(* IEC 61131-3 sources: volt/packages/volt-lsp-iec/test-corpus/pro2193/Device/Plc Logic/Application/09 Misc/Library Manager/AlarmManager (part 3) *)

(* ---- ALARMSTORAGEMANAGER.pou ---- *)
FUNCTION_BLOCK ALARMSTORAGEMANAGER
VAR
	M_ALARMSTORAGE : STI.Storage;
	M_ITFSTORAGE : STO.IStorage;
	M_ITFTABLE : STO.ITable;
	M_ADWROOTPAGES : ARRAY [EAlarmStorageObject.IX_MIN..EAlarmStorageObject.IX_LAST] OF CAA.IDENT;
	M_XROOTPAGESDETERMINED : BOOL;
	M_UDICOUNTLATCHVARIABLES : CAA.COUNT;
	WRITEACCESSNECESSARY : BOOL;
END_VAR
END_FUNCTION_BLOCK

METHOD BEGINTRANSACTION : STO.ITransaction
VAR_INPUT
	XREADONLY : BOOL;
END_VAR
VAR_OUTPUT
	EERROR : STO.ERROR;
END_VAR
END_METHOD

METHOD CLOSETABLE
VAR_INPUT
	ITFTABLE : STO.ITable;
END_VAR
END_METHOD

METHOD ENDTRANSACTION
VAR_INPUT
	ITFTRANSACTION : STO.ITransaction;
	EERROR : STO.ERROR;
END_VAR
END_METHOD

METHOD FB_EXIT : BOOL
VAR_INPUT
	BINCOPYCODE : BOOL;
END_VAR
END_METHOD

METHOD GETCOLUMNIDENTIFIER : CAA.IDENT
VAR_INPUT
	IDCOLUMN : CAA.IDENT;
END_VAR
END_METHOD

METHOD GETNUMBEROFLATCHVARIABLES : CAA.COUNT
VAR_INPUT
	IDBVERSION : INT;
	UDICOUNTCOLUMNSTBLALARM : CAA.COUNT;
END_VAR
END_METHOD

METHOD GETSTORAGE : STO.IStorage
END_METHOD

METHOD OPENTABLE : STO.ITable
VAR_INPUT
	XREADONLY : BOOL;
END_VAR
VAR_OUTPUT
	EERROR : STO.ERROR;
END_VAR
END_METHOD

METHOD DETERMINEROOTPAGES : STO.ERROR
END_METHOD

METHOD GETROOTPAGE : CAA.IDENT
VAR_INPUT
	EDATABASEOBJECT : EAlarmStorageObject;
END_VAR
END_METHOD

METHOD ISREADY : BOOL
END_METHOD

METHOD RESET
END_METHOD

METHOD CLOSESTORAGE
END_METHOD

METHOD DETERMINEROOTPAGESOPENSTORAGE : STO.ERROR
VAR_OUTPUT
	XREOPENREADONLY : BOOL;
END_VAR
END_METHOD

METHOD PRVCHECKJOURNAL
END_METHOD

METHOD PRVHELPGETDATABASEFILEPATH : CAA.FILENAME
END_METHOD

METHOD PRVOPENSTORAGE : STO.ERROR
VAR_INPUT
	XREADONLY : BOOL;
END_VAR
END_METHOD

METHOD PROTCLOSECURSOR : STO.ERROR
VAR_INPUT
	EERRORFROMPREVIOUSPROCESSING : STO.ERROR;
	ICALLINGMETHOD : INT;
END_VAR
VAR_IN_OUT
	ITFCURSOR : STO.ICursor;
END_VAR
END_METHOD

METHOD PROTGETEXCLUSIVETRANSACTION : STO.ITransaction
VAR_INPUT
	ICOUNTRETRIES : INT;
END_VAR
VAR_OUTPUT
	EERROR : STO.ERROR;
END_VAR
END_METHOD

METHOD PROTRELEASEROW : STO.ERROR
VAR_INPUT
	EERRORFROMPREVIOUSPROCESSING : STO.ERROR;
	ICALLINGMETHOD : INT;
END_VAR
VAR_IN_OUT
	ITFROW : STO.IRow;
END_VAR
END_METHOD

(* ---- ALARMSTORAGEQUEUE.pou ---- *)
FUNCTION_BLOCK ALARMSTORAGEQUEUE
VAR
	_PAQUEUE : POINTER TO ARRAY [0..0] OF AlarmStorageRow;
	_IQUEUESIZE : UDINT;
	_INEWESTPOS : UDINT := 0;
	_IOLDESTPOS : UDINT := 0;
	_IITEMCOUNT : UDINT := 0;
	_ALARMSTORAGEROWPROVIDER : AlarmStorageRowProvider;
	_UICOUNTEVENTS : UDINT;
	_PAINITIALQUEUE : POINTER TO AlarmStorageRow;
	_XKEEPOLDVALUES : BOOL;
	_XFIXQUEUENECESSARY : BOOL;
	COUNTALARMSTOINSERT : UDINT;
	COUNTEVENTSTOINSERT : UDINT;
END_VAR
END_FUNCTION_BLOCK

METHOD CANPOSTALARM : BOOL
END_METHOD

METHOD CLEAR
END_METHOD

METHOD FB_EXIT : BOOL
VAR_INPUT
	BINCOPYCODE : BOOL;
END_VAR
END_METHOD

METHOD FB_INIT : BOOL
VAR_INPUT
	BINITRETAINS : BOOL;
	BINCOPYCODE : BOOL;
END_VAR
END_METHOD

METHOD FIXAFTERONLINECHANGEIFNECESSARY
VAR_INPUT
	STORAGE : IDatabaseFileAlarmStorage;
END_VAR
END_METHOD

METHOD GETCURRENTALARM : AlarmStorageRow
END_METHOD

METHOD INIT
VAR_INPUT
	PQUEUEDATA : POINTER TO AlarmStorageRow;
	NUMQUEUEENTRIES : UDINT;
END_VAR
END_METHOD

METHOD ISEMPTY : BOOL
END_METHOD

METHOD ONLINECHANGEDONE
END_METHOD

METHOD ONLINECHANGEPREPARE
END_METHOD

METHOD POSTALARM : BOOL
VAR_INPUT
	ITFALARM : IAlarm;
	ITFDATABASEFILEALARMSTORAGE : IDatabaseFileAlarmStorage;
	ESTATE : AlarmState;
	EPREVSTATE : AlarmState;
	XFORCEUPDATE : BOOL;
END_VAR
VAR_OUTPUT
	ROW : AlarmStorageRow;
END_VAR
END_METHOD

METHOD REMOVECURRENTALARM
END_METHOD

METHOD TRYTOENLARGEQUEUE
END_METHOD

METHOD ASSIGNINITVALUES
END_METHOD

METHOD RESETSTOREDREFERENCES
END_METHOD

METHOD TRYTOENLARGEQUEUEHELP
VAR_INPUT
	KEEPNEWESTPOS : BOOL;
END_VAR
END_METHOD

METHOD PRVGETTYPEDVALUE
VAR_INPUT
	ITFTYPEDVALUE : ITypedValue;
END_VAR
VAR_OUTPUT
	BYTYPECLASS : BYTE;
	LIVALUE : LINT;
END_VAR
END_METHOD

(* ---- ALARMSTORAGEREADER.pou ---- *)
FUNCTION_BLOCK ALARMSTORAGEREADER EXTENDS AlarmStorageManager
VAR_INPUT
	_HLOCK : RTS_IEC_HANDLE := RTS_INVALID_HANDLE;
END_VAR
VAR
	M_DATABASEACCESS : SQLiteDatabaseAccess;
	M_ROWIDITERATOR : AlarmStorageReaderRowIdIterator;
	M_ITFALARMSTORAGEREADERCONSUMER : IAlarmStorageReaderConsumer;
	M_ITFALARMSTORAGEMANAGER : IAlarmStorageManager := THIS^;
	M_EBYTEORDER : EAlarmByteOrder := EAlarmByteOrder.Unknown;
	M_ALATCHVARIABLES : ARRAY [1..2] OF LatchVariable;
	M_AWSLATCHVARVALUE : ARRAY [0..1] OF WSTRING(255);
	M_PALATCHVARSTRINGALLOC : POINTER TO ARRAY [0..10] OF WSTRING(255);
	M_PALATCHVARALLOC : POINTER TO ARRAY [0..10] OF LatchVariable;
	M_ICOUNTLATCHVARALLOC : INT;
	M_LOCKRESULT : RTS_IEC_RESULT;
	M_SWHOHASLOCK : STRING;
END_VAR
END_FUNCTION_BLOCK

METHOD ADDALARMSTORAGELISTENER : EAlarmStorageReaderErrors
VAR_INPUT
	ITFALARMSTORAGELISTENER : IAlarmStorageListener;
END_VAR
END_METHOD

METHOD CONTINUEREADING : EAlarmStorageReaderErrors
VAR_INPUT
	LITIMSTAMPFROM : LINT;
	LITIMSTAMPTO : LINT;
	XREADASCENDING : BOOL;
	ITFALARMSTORAGEREADERCONSUMER : IAlarmStorageReaderConsumer;
END_VAR
END_METHOD

METHOD FB_EXIT : BOOL
VAR_INPUT
	BINCOPYCODE : BOOL;
END_VAR
END_METHOD

METHOD FB_INIT : BOOL
VAR_INPUT
	BINITRETAINS : BOOL;
	BINCOPYCODE : BOOL;
END_VAR
END_METHOD

METHOD GETALARMSFROMSTORAGE : STO.ERROR
VAR_INPUT
	ISKIPROWS : INT;
	IMAXROWS : INT;
	FILTERCRITERIA : REFERENCE TO VisuFbAlarmFilterCriteria;
	ITFALARMDATABLOCK : IAlarmDataBlockBase2;
END_VAR
VAR_IN_OUT
	BROWIDVALID : BOOL;
	DIROWID : DINT;
END_VAR
END_METHOD

METHOD GETALARMSFROMSTORAGE2 : STO.ERROR
VAR_INPUT
	ITFDATABASEACCESS : IDatabaseAccess;
	ISKIPROWS : INT;
	IMAXROWS : INT;
	FILTERCRITERIA : REFERENCE TO VisuFbAlarmFilterCriteria;
	ITFALARMDATABLOCK : IAlarmDataBlockBase2;
END_VAR
VAR_IN_OUT
	BROWIDVALID : BOOL;
	DIROWID : DINT;
END_VAR
END_METHOD

METHOD GETALARMSFROMSTORAGE3 : STO.ERROR
VAR_INPUT
	ITFDATABASEACCESS : IDatabaseAccess3;
	DWROWIDLATEST : DWORD;
	IMAXROWS : INT;
	ITFALARMTRAVERSALCONSUMER : IAlarmTraversalConsumer;
END_VAR
END_METHOD

METHOD GETALARMSFROMSTORAGE4 : STO.ERROR
VAR_INPUT
	ITFDATABASEACCESS : IDatabaseAccess3;
	ITFALARMTRAVERSALCONSUMER : IAlarmTraversalConsumer;
END_VAR
END_METHOD

METHOD GETALARMSFROMSTORAGE5 : STO.ERROR
VAR_INPUT
	DISKIPROWS : DINT;
	DIMAXROWS : DINT;
	FILTERCRITERIA : REFERENCE TO VisuFbAlarmFilterCriteria;
	ITFALARMDATABLOCK : IAlarmDataBlockBase2;
END_VAR
VAR_IN_OUT
	BROWIDVALID : BOOL;
	DIROWID : DINT;
END_VAR
END_METHOD

METHOD GETALARMSFROMSTORAGE6 : STO.ERROR
VAR_INPUT
	ITFDATABASEACCESS : IDatabaseAccess;
	DISKIPROWS : DINT;
	DIMAXROWS : DINT;
	FILTERCRITERIA : REFERENCE TO VisuFbAlarmFilterCriteria;
	ITFALARMDATABLOCK : IAlarmDataBlockBase2;
END_VAR
VAR_IN_OUT
	BROWIDVALID : BOOL;
	DIROWID : DINT;
END_VAR
END_METHOD

METHOD GETCOUNTALARMSFROMSTORAGE : DINT
VAR_INPUT
	FILTERCRITERIA : REFERENCE TO VisuFbAlarmFilterCriteria;
	ITFALARMDATABLOCK : IAlarmDataBlockBase2;
END_VAR
VAR_OUTPUT
	EERROR : STO.ERROR;
	DWCOUNTLATCHVARIABLESINSTORAGE : CAA.COUNT;
END_VAR
END_METHOD

METHOD GETCOUNTALLALARMSFROMSTORAGE : CAA.COUNT
VAR_OUTPUT
	EERROR : STO.ERROR;
END_VAR
END_METHOD

METHOD GETFIRSTLASTROWID : EAlarmStorageReaderErrors
VAR_OUTPUT
	DIROWIDFIRST : DINT;
	DIROWIDLAST : DINT;
END_VAR
END_METHOD

METHOD GETMINMAXTIMESTAMPS : EAlarmStorageReaderErrors
VAR_OUTPUT
	LIMINTIMESTAMP : LINT;
	LIMAXTIMESTAMP : LINT;
	XTABLEISEMPTY : BOOL;
	UDICOUNTALARMS : UDINT;
END_VAR
END_METHOD

METHOD READ : EAlarmStorageReaderErrors
VAR_INPUT
	LITIMSTAMPFROM : LINT;
	LITIMSTAMPTO : LINT;
	XREADASCENDING : BOOL;
	ITFALARMSTORAGEREADERCONSUMER : IAlarmStorageReaderConsumer;
END_VAR
END_METHOD

METHOD REMOVEALARMSTORAGELISTENER : EAlarmStorageReaderErrors
VAR_INPUT
	ITFALARMSTORAGELISTENER : IAlarmStorageListener;
END_VAR
END_METHOD

METHOD SEMAPHOREACQUIRE
VAR_INPUT
	SWHO : STRING;
END_VAR
END_METHOD

METHOD SEMAPHORERELEASE
VAR_INPUT
	SWHO : STRING;
END_VAR
END_METHOD

METHOD PRVALLOCLATCHVARS
VAR_INPUT
	ICNTVAR : INT;
END_VAR
END_METHOD

METHOD PRVDOCONTINUEREADING : BOOL
VAR_INPUT
	DIROWCOUNTER : DINT;
END_VAR
END_METHOD

METHOD PRVFINDROWID : CAA.IDENT
VAR_INPUT
	ITFDATABASEACCESS : IDatabaseAccess;
	XSEARCHFIRST : BOOL;
END_VAR
VAR_OUTPUT
	EERROR : STO.ERROR;
END_VAR
END_METHOD

METHOD PRVFREELATCHVARS
END_METHOD

METHOD PRVREAD : EAlarmStorageReaderErrors
VAR_INPUT
	LITIMSTAMPFROM : LINT;
	LITIMSTAMPTO : LINT;
	XREADASCENDING : BOOL;
END_VAR
END_METHOD

METHOD PRVREADALARMCOMMENT
VAR_INPUT
	IDWHICHCOLUMN : CAA.IDENT;
	ITFDATABASEACCESS4 : IDatabaseAccess4;
END_VAR
VAR_IN_OUT
	EERROR : STO.ERROR;
	CMTBUFFER : AlarmComment;
END_VAR
END_METHOD

METHOD PRVREADLATCHVARSTRING2 : STO.ERROR
VAR_INPUT
	LIROWID : LINT;
	ITFDATABASEACCESS : IDatabaseAccess;
	BYLATCHVARTYPE : BYTE;
	PBVARVALUE : POINTER TO BYTE;
	ISZVARVALUE : INT;
END_VAR
END_METHOD

METHOD PRVREADLATCHVARSTRING : STO.ERROR
VAR_INPUT
	LIROWID : LINT;
	ITFDATABASEACCESS : IDatabaseAccess;
	BYLATCHVARTYPE : BYTE;
END_VAR
VAR_OUTPUT
	CBPSTRING : CharBufferPtr;
END_VAR
END_METHOD

METHOD PRVRETRIEVELATCHVARVALUE : STO.ERROR
VAR_INPUT
	ITFDATABASEACCESS : IDatabaseAccess;
	ITFALARMMETAOBJECTSTUB3 : IAlarmMetaObjectStub3;
	USIWHICHLATCHVAR : USINT;
END_VAR
END_METHOD

METHOD PRVTBLALARMFINDTIMESTAMP : STO.ERROR
VAR_INPUT
	ITFDATABASEACCESS : IDatabaseAccess;
	LITIMSTAMP : LINT;
	XUSENEXTROW : BOOL;
END_VAR
VAR_OUTPUT
	IDROWTIMSTAMP : CAA.IDENT;
END_VAR
END_METHOD

(* ---- ALARMSTORAGEREADERROWIDITERATOR.pou ---- *)
FUNCTION_BLOCK ALARMSTORAGEREADERROWIDITERATOR
VAR
	M_IDROWTBLALARMFROM : CAA.IDENT;
	M_IDROWTBLALARMTO : CAA.IDENT;
	M_IDROWCURR : CAA.IDENT;
	M_XITERATEASCENDING : BOOL;
	M_IDLASTPROCESSEDROWID : CAA.IDENT := AlarmConstants.INVALID_ROWID;
	M_LITIMESTAMP : LINT;
END_VAR
END_FUNCTION_BLOCK

METHOD GETNEXTROWID : CAA.IDENT
END_METHOD

METHOD GETSAVEDSTATE : LINT
END_METHOD

METHOD HASNEXTROWID : BOOL
END_METHOD

METHOD HASSAVEDSTATE : BOOL
END_METHOD

METHOD INITIALIZE
VAR_INPUT
	IDROWTBLALARMFROM : CAA.IDENT;
	IDROWTBLALARMTO : CAA.IDENT;
	XITERATEASCENDING : BOOL;
END_VAR
END_METHOD

METHOD SAVESTATE
VAR_INPUT
	IDLASTPROCESSEDROWID : CAA.IDENT;
	LITIMESTAMP : LINT;
END_VAR
END_METHOD

(* ---- ALARMSTORAGEROW.pou ---- *)
FUNCTION_BLOCK ALARMSTORAGEROW
VAR_INPUT
	UDIALARMID : UDINT;
	UDIALARMCLASSID : UDINT;
	UDIALARMGROUPID : UDINT;
	LITIMESTAPLAST : TIMESTAMP;
	LITIMESTAPACTIVE : TIMESTAMP;
	LITIMESTAPINACTIVE : TIMESTAMP;
	LITIMESTAPACKNOWLEDGE : TIMESTAMP;
	IOFFSETLAST : INT := -1;
	IOFFSETACTIVE : INT := -1;
	IOFFSETINACTIVE : INT := -1;
	IOFFSETACKNOWLEDGE : INT := -1;
	USIPRIORITY : USINT;
	ESTATE : AlarmState;
	EPREVSTATE : AlarmState;
	BYTRIGGERVALUETYPE : BYTE;
	LITRIGGERVALUEVAL : LINT;
	PLATCHVARIABLES : POINTER TO ARRAY [0..10] OF LatchVariable;
	USICOUNTLATCHVARIABLES : USINT;
	ITFALARM : IAlarm;
	ITFDATABASEFILEALARMSTORAGE : IDatabaseFileAlarmStorage;
	IDROW : CAA.IDENT;
	XIDROWVALID : BOOL;
	XFORCEUPDATE : BOOL;
	SREMOTEDEVICENAME : STRING;
	CMTACTIVE : AlarmComment;
	CMTACTIVEACK : AlarmComment;
	CMTWAITINGCONF : AlarmComment;
	CMTNORMAL : AlarmComment;
	XINVALID : BOOL;
END_VAR
END_FUNCTION_BLOCK

METHOD DERIVEALARMREFERENCE
END_METHOD

METHOD GETLATCHVARVALUE
VAR_INPUT
	USIWHICHLATCHVAR : USINT;
END_VAR
VAR_OUTPUT
	BYTYPE : BYTE;
	LIVALUE : LINT;
END_VAR
END_METHOD

METHOD RESETALARMCOMMENTS : BOOL
END_METHOD

METHOD SETLATCHVARVALUE
VAR_INPUT
	USIWHICHLATCHVAR : USINT;
	BYTYPE : BYTE;
	LIVALUE : LINT;
END_VAR
END_METHOD

(* ---- ALARMSTORAGEROWPROVIDER.pou ---- *)
FUNCTION_BLOCK ALARMSTORAGEROWPROVIDER
VAR
	M_PAALARMSTORAGEROWS : POINTER TO ARRAY [0..100] OF AlarmStorageRow;
	M_ICOUNTROWS : UDINT;
	M_PALATCHVARIABLES : POINTER TO ARRAY [0..100] OF LatchVariable;
	M_ICOUNTLATCHVARIABLES : UDINT;
	COMPONENT : STRING := 'AlarmStorageRowProvider';
END_VAR
END_FUNCTION_BLOCK

METHOD ALLOCATEALARMSTORAGEROWARRAY : BOOL
VAR_INPUT
	IREQUIREDARRAYSIZE : UDINT;
	USICOUNTLATCHVARIABLES : USINT;
	PACURRENTQUEUE : POINTER TO AlarmStorageRow;
	ICURRENTQUEUESIZE : UDINT;
	ICURRENTREADINDEX : UDINT;
END_VAR
VAR_OUTPUT
	PANEWQUEUE : POINTER TO ARRAY [0..0] OF AlarmStorageRow;
	INEWQUEUESIZE : UDINT;
END_VAR
END_METHOD

METHOD COPYQUEUECONTENT : BOOL
VAR_INPUT
	PACURRENTQUEUE : POINTER TO AlarmStorageRow;
	ICURRENTQUEUESIZE : UDINT;
	ICURRENTREADINDEX : UDINT;
	PANEWALARMSTORAGEROWS : POINTER TO AlarmStorageRow;
	INEWQUEUESIZE : UDINT;
	PANEWLATCHVARIABLES : POINTER TO LatchVariable;
	USICOUNTLATCHVARIABLES : USINT;
END_VAR
END_METHOD

METHOD FB_EXIT : BOOL
VAR_INPUT
	BINCOPYCODE : BOOL;
END_VAR
END_METHOD

METHOD FREEBUFFER
VAR_INPUT
	PPBYBUFFER : POINTER TO POINTER TO BYTE;
	PICOUNT : POINTER TO INT;
END_VAR
END_METHOD

METHOD FREEBUFFERS
END_METHOD

(* ---- ALLOCATOR.pou ---- *)
FUNCTION_BLOCK ALLOCATOR
VAR_INPUT
	SCOMPONENT : STRING;
END_VAR
VAR
	DITOTMEM : DINT;
	TOTMEM : DINT;
END_VAR
END_FUNCTION_BLOCK

METHOD ALLOCANDCOPYWSTRING : POINTER TO WSTRING
VAR_INPUT
	PWSWHO : POINTER TO WSTRING;
END_VAR
END_METHOD

METHOD ALLOCBYTES : POINTER TO BYTE
VAR_INPUT
	UXISIZE : __UXINT;
	SWHO : STRING;
END_VAR
END_METHOD

METHOD ALLOCPROXYFBALARMCONTAINER : POINTER TO AlarmContainer
VAR_INPUT
	SWHO : STRING;
END_VAR
END_METHOD

METHOD ALLOCPROXYFBALARMMETAOBJECTSTUB : POINTER TO ProxyFbAlarmMetaObjectStub
VAR_INPUT
	SWHO : STRING;
END_VAR
END_METHOD

METHOD ALLOCPROXYSTRUCTALARMCLASSDESCRIPTION : POINTER TO ProxyStructAlarmClass
VAR_INPUT
	SWHO : STRING;
END_VAR
END_METHOD

METHOD ALLOCPROXYSTRUCTALARMDESCRIPTION : POINTER TO ProxyStructAlarm
VAR_INPUT
	SWHO : STRING;
END_VAR
END_METHOD

METHOD ALLOCPROXYSTRUCTALARMGROUPDESCRIPTION : POINTER TO ProxyStructAlarmGroup
VAR_INPUT
	SWHO : STRING;
END_VAR
END_METHOD

METHOD ALLOCPROXYSTRUCTHISTORICALALARMACTIVE : POINTER TO ProxyStructHistoricalAlarmActive
VAR_INPUT
	SWHO : STRING;
END_VAR
END_METHOD

METHOD ALLOCVALUETYPEBUNDLE : POINTER TO ValueTypeBundle
VAR_INPUT
	SWHO : STRING;
END_VAR
END_METHOD

METHOD FREEBYTES
VAR_INPUT
	PTR : POINTER TO BYTE;
	UXISIZE : __UXINT;
END_VAR
END_METHOD

METHOD FREEPROXYFBALARMCONTAINER
VAR_INPUT
	PREQ : POINTER TO AlarmContainer;
END_VAR
END_METHOD

METHOD FREEPROXYFBALARMMETAOBJECTSTUB
VAR_INPUT
	PREQ : POINTER TO ProxyFbAlarmMetaObjectStub;
END_VAR
END_METHOD

METHOD FREEPROXYSTRUCTALARMCLASSDESCRIPTION
VAR_INPUT
	PREQ : POINTER TO ProxyStructAlarmGroup;
END_VAR
END_METHOD

METHOD FREEPROXYSTRUCTALARMDESCRIPTION
VAR_INPUT
	PREQ : POINTER TO ProxyStructAlarm;
END_VAR
END_METHOD

METHOD FREEPROXYSTRUCTALARMGROUPDESCRIPTION
VAR_INPUT
	PREQ : POINTER TO ProxyStructAlarmClass;
END_VAR
END_METHOD

METHOD FREEPROXYSTRUCTHISTORICALALARMACTIVE
VAR_INPUT
	PREQ : POINTER TO ProxyStructHistoricalAlarmActive;
END_VAR
END_METHOD

METHOD FREEVALUETYPEBUNDLE
VAR_INPUT
	PREQ : POINTER TO ValueTypeBundle;
END_VAR
END_METHOD

(* ---- BINTAGWRITERALARMMETAOBJECTSTUB.pou ---- *)
FUNCTION_BLOCK BINTAGWRITERALARMMETAOBJECTSTUB
VAR
	M_ITFTAGGEDSERVICEWRITER : ITaggedServiceWriter;
	M_LITIMESTAMPACKNOWLEDGE : Timestamp;
	M_LITIMESTAMPACTIVE : Timestamp;
	M_LITIMESTAMPINACTIVE : Timestamp;
	M_LITIMESTAMPLAST : Timestamp;
	M_ITFTYPEDVALUETRIGGER : ITypedValue;
	M_IOFFSETACKNOWLEDGE : INT := -1;
	M_IOFFSETACTIVE : INT := -1;
	M_IOFFSETINACTIVE : INT := -1;
	M_IOFFSETLAST : INT := -1;
	M_PALATCHVARIABLES : POINTER TO ARRAY [0..0] OF LatchVariable;
	M_ICOUNTLATCHVARIABLES : INT;
	M_ISTATE : INT;
	M_UDIALARMID : UDINT;
	M_UDIALARMGROUPID : UDINT;
	OFFSETACKNOWLEDGE : INT;
	OFFSETACTIVE : INT;
	OFFSETINACTIVE : INT;
	OFFSETLAST : INT;
END_VAR
END_FUNCTION_BLOCK

METHOD INITIALIZE
VAR_INPUT
	ITFTAGGEDSERVICEWRITER : ITaggedServiceWriter;
END_VAR
END_METHOD

METHOD SETLATCHVARIABLESBUFFER
VAR_INPUT
	PALATCHVARIABLES : POINTER TO ARRAY [0..0] OF LatchVariable;
	ICOUNTLATCHVARIABLES : INT;
END_VAR
END_METHOD

METHOD SETLATCHVAR1VALUE
VAR_INPUT
	ITFTYPEDVALUELATCHVAR1 : ITypedValue;
END_VAR
END_METHOD

METHOD SETLATCHVAR2VALUE
VAR_INPUT
	ITFTYPEDVALUELATCHVAR2 : ITypedValue;
END_VAR
END_METHOD

METHOD SETSTATE
VAR_INPUT
	ISTATE : INT;
END_VAR
END_METHOD

METHOD SETTIMESTAMPACKNOWLEDGE
VAR_INPUT
	LITIMESTAMPACKNOWLEDGE : Timestamp;
END_VAR
END_METHOD

METHOD SETTIMESTAMPACTIVE
VAR_INPUT
	LITIMESTAMPACTIVE : Timestamp;
END_VAR
END_METHOD

METHOD SETTIMESTAMPINACTIVE
VAR_INPUT
	LITIMESTAMPINACTIVE : Timestamp;
END_VAR
END_METHOD

METHOD SETTIMESTAMPLAST
VAR_INPUT
	LITIMESTAMPLAST : Timestamp;
END_VAR
END_METHOD

METHOD SETTRIGGERVALUE
VAR_INPUT
	ITFTYPEDVALUETRIGGER : ITypedValue;
END_VAR
END_METHOD

METHOD GETCOUNTLATCHVARIABLES : USINT
END_METHOD

METHOD GETLATCHVARVALUE : ITypedValue2
VAR_INPUT
	IWHICHLATCHVAR : INT;
END_VAR
END_METHOD

METHOD SETLATCHVARVALUE
VAR_INPUT
	IWHICHLATCHVAR : INT;
	ITFTYPEDVALUELATCHVAR : ITypedValue;
END_VAR
END_METHOD

METHOD SETALARM
VAR_INPUT
	PALARM : POINTER TO Alarm;
END_VAR
END_METHOD

METHOD FILLINGCOMPLETED : UDINT
END_METHOD

METHOD PRVGETTYPE : BYTE
VAR_INPUT
	ITFTYPEDVALUE : ITypedValue;
END_VAR
END_METHOD

METHOD PRVGETVALUE : LWORD
VAR_INPUT
	ITFTYPEDVALUE : ITypedValue;
END_VAR
END_METHOD

METHOD PRVWRITELATCHVARIABLE
VAR_INPUT
	IWHICHLATCHVAR : INT;
END_VAR
END_METHOD

METHOD GETALARMGROUP : STRING
END_METHOD

METHOD GETCHECKSUM : UDINT
END_METHOD

METHOD GETCURRENTVALUE : ITypedValue
END_METHOD

METHOD GETID : ALARM_ID
END_METHOD

METHOD GETLATCHVAR1VALUE : ITypedValue
END_METHOD

METHOD GETLATCHVAR2VALUE : ITypedValue
END_METHOD

METHOD GETSTATE : INT
END_METHOD

METHOD GETTIMESTAMPACKNOWLEDGE : Timestamp
END_METHOD

METHOD GETTIMESTAMPACTIVE : Timestamp
END_METHOD

METHOD GETTIMESTAMPINACTIVE : Timestamp
END_METHOD

METHOD GETTIMESTAMPLAST : Timestamp
END_METHOD

METHOD GETTRIGGERVALUE : ITypedValue
END_METHOD

METHOD SETACKNOWLEDGE
VAR_INPUT
	BACKNOWLEDGEMULTIPLE : BOOL;
END_VAR
END_METHOD

METHOD SETALARMGROUP
VAR_INPUT
	SALARMGROUP : STRING;
END_VAR
END_METHOD

METHOD SETCURRENTLREALVALUE
VAR_INPUT
	LRVALUE : LREAL;
END_VAR
END_METHOD

METHOD SETID
VAR_INPUT
	UIID : ALARM_ID;
END_VAR
END_METHOD

METHOD SWAPVALUES
END_METHOD

METHOD GETALARM : POINTER TO Alarm
END_METHOD

METHOD SETCURRENTVALUE
VAR_INPUT
	ITFTYPEDVALUECURRENT : ITypedValue;
END_VAR
END_METHOD

(* ---- BINTAGWRITERDATABLOCK.pou ---- *)
FUNCTION_BLOCK BINTAGWRITERDATABLOCK
VAR
	M_BINTAGWRITERALARMMETAOBJECTSTUB : BinTagWriterAlarmMetaObjectStub;
	M_ICOUNTROWS : INT;
END_VAR
END_FUNCTION_BLOCK

METHOD GETALARMMETAOBJECTSTUB : IAlarmMetaObjectStub3
VAR_INPUT
	IROW : INT;
	IOFFSET : INT;
END_VAR
END_METHOD

METHOD GETCOUNTROWS : INT
END_METHOD

METHOD INITIALIZE
VAR_INPUT
	ITFTAGGEDSERVICEWRITER : ITaggedServiceWriter;
END_VAR
END_METHOD

METHOD SETCOUNTROWS : BOOL
VAR_INPUT
	ICOUNT : INT;
END_VAR
END_METHOD

METHOD SETLATCHVARIABLESBUFFER
VAR_INPUT
	PALATCHVARIABLES : POINTER TO ARRAY [0..0] OF LatchVariable;
	ICOUNTLATCHVARIABLES : INT;
END_VAR
END_METHOD

METHOD HASALARMS : BOOL
END_METHOD

METHOD SETTOTALCOUNTROWS : BOOL
VAR_INPUT
	DICOUNT : DINT;
END_VAR
END_METHOD

(* ---- CHANGEOBSERVATIONTYPE.pou ---- *)
FUNCTION_BLOCK CHANGEOBSERVATIONTYPE
VAR_INPUT
	M_UIID : ALARM_ID;
	M_ITFCHANGEEVALUATOR : IChangeEvaluator;
END_VAR
END_FUNCTION_BLOCK

METHOD ISACTIVE : BOOL
VAR_INPUT
	ECURRSTATE : AlarmState;
END_VAR
END_METHOD

METHOD ISIMMEDIATELYACTIVE : BOOL
END_METHOD

(* ---- COMMENTCOMPARER.pou ---- *)
FUNCTION_BLOCK COMMENTCOMPARER EXTENDS TSLastComparer
END_FUNCTION_BLOCK

METHOD COMPARE : INT
VAR_INPUT
	DIINDEXALARM1 : DINT;
	DIINDEXALARM2 : DINT;
END_VAR
END_METHOD

(* ---- COMPONENTREGISTRATOR.pou ---- *)
FUNCTION_BLOCK COMPONENTREGISTRATOR
VAR
	_HCOMPONENT : RTS_IEC_HANDLE;
	CMINVALIDHANDLE : RTS_IEC_HANDLE := 16#FFFFFFFF;
END_VAR
END_FUNCTION_BLOCK

METHOD FB_EXIT : BOOL
VAR_INPUT
	BINCOPYCODE : BOOL;
END_VAR
END_METHOD

METHOD FB_INIT
VAR_INPUT
	BINITRETAINS : BOOL;
	BINCOPYCODE : BOOL;
END_VAR
END_METHOD

(* ---- CONVERTIECTYPEDLITERAL.pou ---- *)
FUNCTION_BLOCK CONVERTIECTYPEDLITERAL
VAR
	CH_PLUS : BYTE := 16#2B;
	CH_MINUS : BYTE := 16#2D;
	CH_POINT : BYTE := 16#2E;
	CH_0 : BYTE := 16#30;
	CH_1 : BYTE := 16#31;
	CH_2 : BYTE := 16#32;
	CH_3 : BYTE := 16#33;
	CH_4 : BYTE := 16#34;
	CH_5 : BYTE := 16#35;
	CH_6 : BYTE := 16#36;
	CH_7 : BYTE := 16#37;
	CH_8 : BYTE := 16#38;
	CH_9 : BYTE := 16#39;
	CH_COLON : BYTE := 16#3A;
	CH_A : BYTE := 16#41;
	CH_B : BYTE := 16#42;
	CH_C : BYTE := 16#43;
	CH_D : BYTE := 16#44;
	CH_E : BYTE := 16#45;
	CH_F : BYTE := 16#46;
	CH_H : BYTE := 16#48;
	CH_M : BYTE := 16#4D;
	CH_N : BYTE := 16#4E;
	CH_S : BYTE := 16#53;
	CH_U : BYTE := 16#55;
END_VAR
END_FUNCTION_BLOCK

METHOD CONVERT : INT
VAR_INPUT
	SLITERAL : STRING(255);
	XCONVERTCHECK : BOOL;
END_VAR
VAR_OUTPUT
	VTYPE : Visu_Types;
	LIVALUE : LINT;
	RVALUE : REAL;
	LRVALUE : LREAL;
END_VAR
END_METHOD

METHOD TEST : STRING
END_METHOD

METHOD CONVERTOLD : INT
VAR_INPUT
	PLITERAL : POINTER TO STRING(255);
END_VAR
VAR_OUTPUT
	VTYPE : Visu_Types;
	LIVALUE : LINT;
	RVALUE : REAL;
	LRVALUE : LREAL;
END_VAR
END_METHOD

METHOD PRVANALYSEDURATIONVALUE : LINT
VAR_INPUT
	PNUMBER : POINTER TO STRING(255);
	LIUNIT : LINT;
END_VAR
END_METHOD

METHOD PRVGETDATE : BOOL
VAR_INPUT
	PTOKEN : POINTER TO STRING(255);
END_VAR
VAR_OUTPUT
	LIDATE : LINT;
END_VAR
END_METHOD

METHOD PRVGETDATEANDTIME : BOOL
VAR_INPUT
	PTOKEN : POINTER TO STRING(255);
END_VAR
VAR_OUTPUT
	LIDT : LINT;
END_VAR
END_METHOD

METHOD PRVGETDURATION : BOOL
VAR_INPUT
	PTOKEN : POINTER TO STRING(255);
END_VAR
VAR_OUTPUT
	LIDURATION : LINT;
END_VAR
END_METHOD

METHOD PRVGETFACTOR
VAR_INPUT
	LIBASE : LINT;
	PSUB : POINTER TO STRING;
END_VAR
VAR_OUTPUT
	LIFACTOR : LINT;
END_VAR
END_METHOD

METHOD PRVGETLREAL : BOOL
VAR_INPUT
	PTOKEN : POINTER TO STRING(255);
END_VAR
VAR_OUTPUT
	LRVALUE : LREAL;
END_VAR
END_METHOD

METHOD PRVGETNUMERICAL : BOOL
VAR_INPUT
	PTOKEN : POINTER TO STRING(255);
	XSIGNALLOWED : BOOL;
END_VAR
VAR_OUTPUT
	LIVALUE : LINT;
	SBASE16VALUE : STRING;
END_VAR
END_METHOD

METHOD PRVGETREAL : BOOL
VAR_INPUT
	PTOKEN : POINTER TO STRING(255);
END_VAR
VAR_OUTPUT
	RVALUE : REAL;
END_VAR
END_METHOD

METHOD PRVGETTIMEOFDAY : BOOL
VAR_INPUT
	PTOKEN : POINTER TO STRING(255);
END_VAR
VAR_OUTPUT
	LITOD : LINT;
END_VAR
END_METHOD

METHOD PRVINTTODATE : BOOL
VAR_INPUT
	IDAY : INT;
	IMONTH : INT;
	IYEAR : INT;
END_VAR
VAR_OUTPUT
	UIDAYS : UINT;
END_VAR
END_METHOD

METHOD PRVSPLIT
VAR_INPUT
	PSTRING : POINTER TO STRING(255);
	SSPLITCHAR : STRING;
END_VAR
VAR_OUTPUT
	SLEFT : STRING(255);
	SRIGHT : STRING(255);
END_VAR
END_METHOD

(* ---- DATABASEACCESSERRORHANDLER.pou ---- *)
FUNCTION_BLOCK DATABASEACCESSERRORHANDLER
VAR_INPUT
	M_UIDISKFULLDATABASEACCESSSUSPENDTIME : UINT;
END_VAR
VAR
	M_XLOGERRORS : BOOL := TRUE;
	M_XDATABASEACCESSENABLED : BOOL := TRUE;
	M_DWTIMESTAMPFIRSTDISKFULLEVENT : DWORD;
END_VAR
END_FUNCTION_BLOCK

METHOD ERRORHANDLING
VAR_INPUT
	IFUNCTION : INT;
	IERRCODE : INT;
END_VAR
END_METHOD

METHOD ISDATABASEACCESSENABLED : BOOL
END_METHOD

METHOD ISSEARCHNOTFOUNDERROR : BOOL
VAR_INPUT
	EERROR : STO.ERROR;
END_VAR
END_METHOD

METHOD SQLITEERRORHANDLING
VAR_INPUT
	IFUNCTION : INT;
	EERROR : STO.ERROR;
	IACTION : INT;
END_VAR
END_METHOD

METHOD SQLITEERRORHANDLINGSEARCHING
VAR_INPUT
	IFUNCTION : INT;
	EERROR : STO.ERROR;
	IACTION : INT;
END_VAR
END_METHOD

METHOD PRVGETFUNCTIONNAME : STRING
VAR_INPUT
	IFUNCTION : INT;
END_VAR
END_METHOD

(* ---- DATABASEFILEALARMSTORAGE.pou ---- *)
FUNCTION_BLOCK DATABASEFILEALARMSTORAGE EXTENDS AlarmStorageManager
VAR
	M_SAPPLICATIONNAME : STRING;
	M_AITFALARMSTORAGELISTENER : ARRAY [0..(COUNT_MAX_ALARM_STORAGE_LISTENER - 1)] OF IAlarmStorageListener;
	M_SOLDREMOTEDEVICENAME : STRING;
	M_LIREMOTEDEVICENAMEVALUE : LINT;
	M_CACHEDDBVERSION : INT := UNDETERMINED_DB_VERSION;
	M_CACHEDDBVERSIONERROR : STO.ERROR;
	M_WRITECONTEXT : DatabaseFileWriteContext;
	M_XCHANGESTATETONORMAL : BOOL;
	M_XASSIGNINACTIVETIMESTAMPS : BOOL;
	COUNT_MAX_ALARM_STORAGE_LISTENER : INT := 5;
	UNDETERMINED_DB_VERSION : INT := -1;
	ASSIGNINACTIVETIMESTAMPS : BOOL;
	CHANGESTATETONORMAL : BOOL;
	TABLE : STO.ITable;
	WRITEACCESSNECESSARY : BOOL;
END_VAR
END_FUNCTION_BLOCK

METHOD GETDATABASEFILEPATH : STRING
END_METHOD

METHOD GETFILELIMIT : FileLimit
END_METHOD

METHOD GETMAXRECORDCOUNT : UDINT
END_METHOD

METHOD GETSUBDIRECTORY : STRING
END_METHOD

METHOD WRITETOSTORAGE : STO.ERROR
VAR_INPUT
	ITFTABLE : STO.ITable;
	ROW : AlarmStorageRow;
	ICOUNTRETRIES : INT;
END_VAR
END_METHOD

METHOD CLEARBUFFER
END_METHOD

METHOD ADDALARMSTORAGELISTENER : EAlarmStorageReaderErrors
VAR_INPUT
	ITFALARMSTORAGELISTENER : IAlarmStorageListener;
END_VAR
END_METHOD

METHOD CREATEALARMSTORAGEMETADATAFILE
VAR_INPUT
	UDICOUNTCOLUMNSTBLALARM : CAA.COUNT;
END_VAR
END_METHOD

METHOD OPENTABLE2 : STO.ITable
VAR_INPUT
	XREADONLY : BOOL;
END_VAR
VAR_OUTPUT
	EERROR : STO.ERROR;
END_VAR
END_METHOD

METHOD REMOVEALARMSTORAGELISTENER : EAlarmStorageReaderErrors
VAR_INPUT
	ITFALARMSTORAGELISTENER : IAlarmStorageListener;
END_VAR
END_METHOD

METHOD CHECKFILELIMITREACHED : STO.Error
VAR_INPUT
	ITFTABLE : STO.ITable;
	ICOUNTRETRIES : INT;
	ICOUNTROWSTOINSERT : INT;
END_VAR
END_METHOD

METHOD GETEXCLUSIVETRANSACTION : STO.ITransaction
VAR_INPUT
	ICOUNTRETRIES : INT;
END_VAR
VAR_OUTPUT
	EERROR : STO.ERROR;
END_VAR
END_METHOD

METHOD WRITETOSTORAGE2 : STO.ERROR
VAR_INPUT
	ITFTABLE : STO.ITable;
	ROW : AlarmStorageRow;
	ITFTRANSACTION : STO.ITransaction;
END_VAR
END_METHOD

METHOD DELETEALARMSTORAGEFILE : STO.ERROR
VAR_INPUT
	SFILEPATH : CAA.FILENAME;
END_VAR
END_METHOD

METHOD GETALARMSFROMSTORAGE : STO.ERROR
VAR_INPUT
	ISKIPROWS : INT;
	IMAXROWS : INT;
	FILTERCRITERIA : REFERENCE TO VisuFbAlarmFilterCriteria;
	ITFALARMDATABLOCK : IAlarmDataBlockBase2;
END_VAR
VAR_IN_OUT
	BROWIDVALID : BOOL;
	DIROWID : DINT;
END_VAR
END_METHOD

METHOD GETCOUNTALARMSFROMSTORAGE : DINT
VAR_INPUT
	FILTERCRITERIA : REFERENCE TO VisuFbAlarmFilterCriteria;
	ITFALARMDATABLOCK : IAlarmDataBlockBase2;
END_VAR
VAR_OUTPUT
	EERROR : STO.ERROR;
	DWCOUNTLATCHVARIABLESINSTORAGE : CAA.COUNT;
END_VAR
END_METHOD

METHOD CREATEWRITECONTEXT : IDatabaseFileWriteContext
END_METHOD

METHOD SCANSTORAGE : STO.ERROR
VAR_INPUT
	ITFCONSUMER : IRemoteDeviceTraversalConsumer;
END_VAR
VAR_OUTPUT
	IVERSION : INT;
	DIREMOTEENTRIESCNT : DINT;
END_VAR
END_METHOD

METHOD WRITETOSTORAGE3 : STO.ERROR
VAR_INPUT
	WRITECONTEXT : IDatabaseFileWriteContext;
	ROW : AlarmStorageRow;
	XFORCEINSERT : BOOL;
	XFIRST : BOOL;
END_VAR
END_METHOD

METHOD CLEARALARMSINSTATENORMAL : STO.Error
VAR_INPUT
	ITFTABLE : STO.ITable;
END_VAR
VAR_OUTPUT
	XFINISHED : BOOL;
END_VAR
VAR_IN_OUT
	DIREMAININGROWCOUNT : DINT;
END_VAR
END_METHOD

METHOD ROWSELECT : STO.IRow
VAR_INPUT
	ITFTABLE : STO.ITable;
	IDROW : CAA.IDENT;
END_VAR
END_METHOD

METHOD CHECKRECORDLIMITREACHED : STO.Error
VAR_INPUT
	ITFTABLE : STO.ITable;
	ICOUNTRETRIES : INT;
	ICOUNTROWSTOINSERT : INT;
	XFORCE : BOOL;
END_VAR
VAR_OUTPUT
	XLIMIT : BOOL;
	UDIMAXRECORDCOUNT : UDINT;
END_VAR
END_METHOD

METHOD DELETEALARMS : STO.Error
VAR_INPUT
	ITFTABLE : STO.ITable;
	ICOUNTRETRIES : INT;
	DICOUNTROWSTODELETE : DINT;
END_VAR
VAR_OUTPUT
	DIROWSDELETED : DINT;
END_VAR
END_METHOD

METHOD GETRECORDSIZE : INT
END_METHOD

METHOD GETSTORAGESIZE : LINT
END_METHOD

METHOD SETEMPTYTIMESTAMPINACTIVETOSTARTTIME : STO.Error
VAR_INPUT
	ITFTABLE : STO.ITable;
END_VAR
END_METHOD

METHOD CHECKFILELIMITREACHEDUDINT : STO.ERROR
VAR_INPUT
	ITFTABLE : STO.ITable;
	ICOUNTRETRIES : INT;
	UDICOUNTROWSTOINSERT : UDINT;
END_VAR
END_METHOD

METHOD CHECKRECORDLIMITREACHEDUDINT : STO.ERROR
VAR_INPUT
	ITFTABLE : STO.ITable;
	ICOUNTRETRIES : INT;
	UDICOUNTROWSTOINSERT : UDINT;
	XFORCE : BOOL;
END_VAR
VAR_OUTPUT
	XLIMIT : BOOL;
	UDIMAXRECORDCOUNT : UDINT;
END_VAR
END_METHOD

METHOD PRVCHECKFILELIMITREACHED : STO.Error
VAR_INPUT
	ITFTABLE : STO.ITable;
	ICOUNTRETRIES : INT;
	UDICOUNTROWSTOINSERT : UDINT;
END_VAR
END_METHOD

METHOD PRVCHECKRECORDLIMITREACHED : STO.Error
VAR_INPUT
	ITFTABLE : STO.ITable;
	ICOUNTRETRIES : INT;
	UDICOUNTROWSTOINSERT : UDINT;
	XFORCE : BOOL;
END_VAR
VAR_OUTPUT
	XLIMIT : BOOL;
	UDIMAXRECORDCOUNT : UDINT;
END_VAR
END_METHOD

METHOD PRVDELETEALARMSTOREACHLIMIT : BOOL
VAR_INPUT
	ITFTABLE : STO.ITable;
	ICOUNTRETRIES : INT;
	UDICOUNTROWSTODELETE : UDINT;
END_VAR
VAR_OUTPUT
	IROWSDELETED : INT;
	EERROR : STO.ERROR;
END_VAR
END_METHOD

METHOD PRVFINDLATCHVARSTRING
VAR_INPUT
	CBPINPUTSTRING : CharBufferPtr;
	BYTYPECLASS : BYTE;
	IVERSION : INT;
	ITFTABLE : STO.ITable;
END_VAR
VAR_OUTPUT
	DIROWID : DINT;
	XFOUND : BOOL;
END_VAR
VAR_IN_OUT
	EERROR : STO.ERROR;
	WSINPUTSTRING : WSTRING(255);
END_VAR
END_METHOD

METHOD PRVFINDLATCHVARSTRING_DBVERBEFORE5
VAR_INPUT
	CBPINPUTSTRING : CharBufferPtr;
	BYTYPECLASS : BYTE;
	ITFCURSOR : STO.ICursor;
END_VAR
VAR_OUTPUT
	DIROWID : DINT;
	XFOUND : BOOL;
END_VAR
VAR_IN_OUT
	EERROR : STO.ERROR;
END_VAR
END_METHOD

METHOD PRVFINDLATCHVARSTRING_DBVERRECENT
VAR_INPUT
	ITFCURSOR : STO.ICursor;
END_VAR
VAR_OUTPUT
	DIROWID : DINT;
	XFOUND : BOOL;
END_VAR
VAR_IN_OUT
	EERROR : STO.ERROR;
	WSINPUTSTRING : WSTRING(255);
END_VAR
END_METHOD

METHOD PRVGETDATABASEFILEPATH : STRING
VAR_INPUT
	SVERSIONINCOMPATIBLECHANGE : STRING;
END_VAR
VAR_OUTPUT
	EERROR : STO.ERROR;
END_VAR
END_METHOD

METHOD PRVGETVERSION : STO.ERROR
VAR_OUTPUT
	IVERSION : INT;
END_VAR
END_METHOD

METHOD PRVGETVERSIONFROMDATABASE : STO.ERROR
VAR_OUTPUT
	IVERSION : INT;
END_VAR
END_METHOD

METHOD PRVREMOVERECORDLIMITREACHED : STO.Error
VAR_INPUT
	UDIMAXRECORDCOUNT : UDINT;
	ITFTABLE : STO.ITable;
	ICOUNTRETRIES : INT;
	ICOUNTROWSTOINSERT : UDINT;
END_VAR
END_METHOD

METHOD PRVSEARCHMINROWIDS : STO.ERROR
VAR_INPUT
	ITFTABLE : STO.ITable;
	ICOUNTROWSIDSTOSEARCH : INT;
	PADWROWIDS : POINTER TO ARRAY [0..50] OF CAA.IDENT;
	IEFFECTIVEARRAYSIZE : INT;
END_VAR
VAR_OUTPUT
	ICOUNTROWSIDS : INT;
END_VAR
END_METHOD

METHOD PRVSETTYPEDVALUE : STO.ERROR
VAR_INPUT
	BYTYPECLASS : BYTE;
	LIVALUE : LINT;
	ITFROWBASE : STO.IRowBase;
	COLVALUE : CAA.IDENT;
	COLTYPE : CAA.IDENT;
END_VAR
END_METHOD

METHOD PRVSORTROWIDS
VAR_INPUT
	PADWROWIDS : POINTER TO ARRAY [0..0] OF CAA.IDENT;
	NFIRST : INT;
	NLAST : INT;
END_VAR
END_METHOD

METHOD PRVSTOREALARMCOMMENTS : STO.ERROR
VAR_INPUT
	PROW : POINTER TO AlarmStorageRow;
	ITFROWPLANCHET : STO.IRowPlanchet;
	ITFROW : STO.IRow;
END_VAR
END_METHOD

METHOD PRVUPDATEROW : BOOL
VAR_INPUT
	HTASK : RTS_IEC_HANDLE;
	ITFROW : STO.IRow;
	ICOUNTRETRIES : INT;
	EERROR : STO.ERROR;
END_VAR
END_METHOD

METHOD PRVWRITEALARMCOMMENTCOLUMN
VAR_INPUT
	PWSVALUE : POINTER TO WSTRING;
	ITFROWPLANCHET : STO.IRowPlanchet;
	ITFROW : STO.IRow;
	DATABASEIDENT : CAA.IDENT;
	ERRACTION : INT;
END_VAR
VAR_IN_OUT
	EERROR : STO.ERROR;
END_VAR
END_METHOD

METHOD PRVWRITEBYTEORDERFLAG
END_METHOD

METHOD PRVWRITELATCHVARSTRINGS
VAR_INPUT
	ITFROWBASE : STO.IRowBase;
	PROW : POINTER TO AlarmStorageRow;
	WRITECONTEXT : IDatabaseFileWriteContext;
END_VAR
VAR_IN_OUT
	EERROR : STO.ERROR;
END_VAR
END_METHOD

METHOD PRVWRITETOSTORAGE : STO.ERROR
VAR_INPUT
	WRITECONTEXT : IDatabaseFileWriteContext;
	ROW : AlarmStorageRow;
	ICOUNTRETRIES : INT;
	XCHECKFILELIMITREACHED : BOOL;
	XFORCEINSERT : BOOL;
END_VAR
END_METHOD

METHOD PRVWRITETOTBLLATCHVARSTRINGS : STO.ERROR
VAR_INPUT
	WRITECONTEXT : IDatabaseFileWriteContext;
	CBPINPUTSTRING : CharBufferPtr;
	BYTYPECLASS : BYTE;
END_VAR
VAR_OUTPUT
	DIROWID : DINT;
END_VAR
END_METHOD

METHOD PRVWRITETRIGGERVALUE
VAR_INPUT
	ITFROWBASE : STO.IRowBase;
	BYTRIGGERVALUETYPE : BYTE;
	LITRIGGERVALUEVAL : LINT;
END_VAR
VAR_IN_OUT
	EERROR : STO.ERROR;
END_VAR
END_METHOD

(* ---- DATABASEFILEWRITECONTEXT.pou ---- *)
FUNCTION_BLOCK DATABASEFILEWRITECONTEXT EXTENDS DatabaseFileWriteContextBase
VAR
	_INUSE : BOOL;
	M_ICOUNTRETRIES : INT := AlarmConstants.RETRY_COUNT;
	M_ICOUNTCYCLEWAIT : INT;
END_VAR
END_FUNCTION_BLOCK

METHOD INITIALIZE : BOOL
VAR_IN_OUT
	DB : DatabaseFileAlarmStorage;
END_VAR
END_METHOD

METHOD RELEASE
VAR_INPUT
	EERRORFORCOMMIT : STO.ERROR;
END_VAR
END_METHOD

METHOD PRVINCREASERETRYCOUNT : BOOL
END_METHOD

METHOD PRVRESETRETRYCOUNT : BOOL
END_METHOD

(* ---- DATABASEFILEWRITECONTEXTBASE.pou ---- *)
FUNCTION_BLOCK DATABASEFILEWRITECONTEXTBASE
VAR
	_MAINTABLE : STO.ITable;
	_STRINGLATCHTABLE : STO.ITable;
	_TRANSACTION : STO.ITransaction;
	_STORAGEMAN : REFERENCE TO DatabaseFileAlarmStorage;
	MAINTABLE : STO.ITable;
	TRANSACTION : STO.ITransaction;
END_VAR
END_FUNCTION_BLOCK

METHOD GETSTRINGLATCHTABLE : STO.ITable
VAR_OUTPUT
	EERROR : STO.ERROR;
END_VAR
END_METHOD

METHOD RELEASE
VAR_INPUT
	EERRORFORCOMMIT : STO.ERROR;
END_VAR
END_METHOD

(* ---- DATABASEFILEWRITECONTEXTTEMPORARY.pou ---- *)
FUNCTION_BLOCK DATABASEFILEWRITECONTEXTTEMPORARY EXTENDS DatabaseFileWriteContextBase
END_FUNCTION_BLOCK

METHOD FB_EXIT : BOOL
VAR_INPUT
	BINCOPYCODE : BOOL;
END_VAR
END_METHOD

METHOD INITIALIZE : BOOL
VAR_INPUT
	MAINTABLE : STO.ITable;
	TRANSACTION : STO.ITransaction;
END_VAR
VAR_IN_OUT
	STORAGEMAN : DatabaseFileAlarmStorage;
END_VAR
END_METHOD

(* ---- DATABASESIZELIMIT.pou ---- *)
FUNCTION_BLOCK DATABASESIZELIMIT
VAR
	M_XINITIALIZED : BOOL;
	M_XFIRST : BOOL := TRUE;
	M_XFIRSTREMOVE : BOOL := TRUE;
	M_METRICS : STO.METRICS;
	M_ITFDATABASEFILEALARMSTORAGE7 : IDatabaseFileAlarmStorage7;
	M_ITFALARMSTORAGEMANAGER : IAlarmStorageManager;
	M_SYSRECORDSIZE : INT;
	M_LISTORAGESIZE : LINT;
	M_XERRORDISPLAYED : BOOL;
	M_LIFILESIZEINERROR : LINT;
	M_ICNTREORGERR : INT;
	M_XBLOCKED : BOOL;
	M_ITEMPREDUCTIONRECORDNUM : INT;
	M_TLASTREORGTIME : TIME;
	M_ICNTDBREORD : INT;
	ISBLOCKED : BOOL;
	LASTREORDERINGTIME : TIME;
	REORDERINGCOUNT : INT;
END_VAR
END_FUNCTION_BLOCK

METHOD CHECKFORSIZELIMIT : BOOL
END_METHOD

METHOD INITIALIZE
VAR_INPUT
	ITFDATABASEFILEALARMSTORAGE : IDatabaseFileAlarmStorage;
END_VAR
END_METHOD

METHOD PRVDBMETRICS : STO.ERROR
VAR_OUTPUT
	MMETRICS : STO.METRICS;
END_VAR
END_METHOD

METHOD PRVGETRECORDSIZE : INT
END_METHOD

METHOD PRVGETRECORDSTOREMOVE : DINT
VAR_INPUT
	LIBYTESTOREMOVE : LINT;
END_VAR
VAR_OUTPUT
	IRECORDSIZE : INT;
END_VAR
END_METHOD

METHOD PRVREORGDB : STO.ERROR
END_METHOD

(* ---- DEFAULTALARMFILTERCRITERIA.pou ---- *)
FUNCTION_BLOCK DEFAULTALARMFILTERCRITERIA
END_FUNCTION_BLOCK

METHOD AREALLALARMCLASSESSELECTED : BOOL
END_METHOD

METHOD AREALLALARMGROUPSSELECTED : BOOL
END_METHOD

METHOD GETALARMCLASSES : POINTER TO ARRAY [0..0] OF UDINT
END_METHOD

METHOD GETALARMGROUPS : POINTER TO ARRAY [0..0] OF UDINT
END_METHOD

METHOD GETCOUNTALARMCLASSES : INT
END_METHOD

METHOD GETCOUNTALARMGROUPS : INT
END_METHOD

METHOD GETPRIORITYFROM : USINT
END_METHOD

METHOD GETPRIORITYTO : USINT
END_METHOD

(* ---- EVENTDISPATCHER.pou ---- *)
FUNCTION_BLOCK EVENTDISPATCHER
VAR
	_HGETCOUNTEVENT : RTS_IEC_HANDLE := Events.Invalid_Handle;
	_HGETCOUNTEVENTINTERFACE : RTS_IEC_HANDLE := Events.Invalid_Handle;
	_HGETALARMSEVENT : RTS_IEC_HANDLE := Events.Invalid_Handle;
	_HGETALARMSEVENTINTERFACE : RTS_IEC_HANDLE := Events.Invalid_Handle;
	_HCHANNELCLOSEDEVENT : RTS_IEC_HANDLE := Events.Invalid_Handle;
	_HCHANNELCLOSEDEVENTINTERFACE : RTS_IEC_HANDLE := Events.Invalid_Handle;
	_HHANDLESERVICEEVENT : RTS_IEC_HANDLE := Events.Invalid_Handle;
	_HHANDLESERVICEEVENTINTERFACE : RTS_IEC_HANDLE := Events.Invalid_Handle;
	_SERVICEHANDLER : AlarmServiceHandler;
END_VAR
END_FUNCTION_BLOCK

METHOD EVENTCALLBACK : UDINT
VAR_INPUT
	PEVENTPARAM : POINTER TO EventParam;
END_VAR
END_METHOD

METHOD FB_EXIT : BOOL
VAR_INPUT
	BINCOPYCODE : BOOL;
END_VAR
END_METHOD

METHOD FB_INIT : BOOL
VAR_INPUT
	BINITRETAINS : BOOL;
	BINCOPYCODE : BOOL;
END_VAR
END_METHOD

(* ---- EXPRESSIONOBSERVATIONTYPE.pou ---- *)
FUNCTION_BLOCK EXPRESSIONOBSERVATIONTYPE
VAR_INPUT
	M_UIID : ALARM_ID;
	M_EXPRESSIONEVALUATOR : IExpressionEvaluator;
END_VAR
END_FUNCTION_BLOCK

METHOD ISACTIVE : BOOL
VAR_INPUT
	ECURRSTATE : AlarmState;
END_VAR
END_METHOD

METHOD ISIMMEDIATELYACTIVE : BOOL
END_METHOD

(* ---- FORMATSTRINGSCANNER.pou ---- *)
FUNCTION_BLOCK FORMATSTRINGSCANNER
END_FUNCTION_BLOCK

METHOD GETFORMATSTRING : BOOL
VAR_INPUT
	RCBSMESSAGE : REFERENCE TO CharBufferString;
	PCBSPLACEHOLDER : POINTER TO CharBufferString;
	IOFFSET : INT;
	ILENGTHPREFIX : INT;
END_VAR
VAR_OUTPUT
	SFORMATSTRING : STRING;
	ITOTALPLACEHOLDERLENGTH : INT;
END_VAR
END_METHOD

(* ---- HASHTABLEKEYELEMENT.pou ---- *)
FUNCTION_BLOCK HASHTABLEKEYELEMENT EXTENDS InstanceBase
VAR
	_INSTANCEPOINTER : POINTER TO BYTE;
	_ALARMTEMPLATENAME : POINTER TO STRING;
	_LIHASH : LINT;
	ALARMTEMPLATENAME : POINTER TO STRING;
	INSTANCEPOINTER : POINTER TO BYTE;
END_VAR
END_FUNCTION_BLOCK

METHOD ELEMENTCOMPARETO : INT
VAR_INPUT
	ITFELEMENT : COL.IElement;
END_VAR
END_METHOD

METHOD ELEMENTEQUALS : BOOL
VAR_INPUT
	ITFELEMENT : COL.IElement;
END_VAR
END_METHOD

METHOD ELEMENTHASHCODE : LINT
END_METHOD

METHOD PRVCALCULATEHASH : LINT
END_METHOD

METHOD PRVINSTINIT : COL.FBF.ERROR
VAR_INPUT
	ITFDATA : COL.FBF.IData;
END_VAR
END_METHOD

(* ---- HASHTABLEKEYELEMENTDATA.pou ---- *)
FUNCTION_BLOCK HASHTABLEKEYELEMENTDATA EXTENDS InstanceData
VAR_INPUT
	PALARMINSTANCE : POINTER TO BYTE;
	STALARMTEMPLATENAME : POINTER TO STRING;
END_VAR
END_FUNCTION_BLOCK

(* ---- HASHTABLEKEYELEMENTFACTORY.pou ---- *)
FUNCTION_BLOCK HASHTABLEKEYELEMENTFACTORY EXTENDS FactoryBase
VAR
	PRVINSTCOUNT : CAA.COUNT;
	PRVINSTPOOLEXTENDSFACTOR : USINT;
	PRVINSTSIZE : CAA.SIZE;
END_VAR
END_FUNCTION_BLOCK

METHOD CREATE : IHashtableKeyElement
VAR_INPUT
	INSTANCEPOINTER : POINTER TO BYTE;
	PSTALARMTEMPLATENAME : POINTER TO STRING;
END_VAR
VAR_OUTPUT
	EERROR : COL.FBF.ERROR;
END_VAR
END_METHOD

(* ---- HASHTABLEVALUEELEMENT.pou ---- *)
FUNCTION_BLOCK HASHTABLEVALUEELEMENT EXTENDS InstanceBase
VAR
	_UDIALARMGROUPID : UDINT;
	_UITEMPLATEALARMSOFFSET : UINT;
	_UITEMPLATEALARMSLENGTH : UINT;
	_UITEMPLATEEVENTSOFFSET : UINT;
	_UITEMPLATEEVENTSLENGTH : UINT;
	ALARMGROUPID : UDINT;
	TEMPLATEALARMSLENGTH : UINT;
	TEMPLATEALARMSOFFSET : UINT;
	TEMPLATEEVENTSLENGTH : UINT;
	TEMPLATEEVENTSOFFSET : UINT;
END_VAR
END_FUNCTION_BLOCK

METHOD ELEMENTCOMPARETO : INT
VAR_INPUT
	ITFELEMENT : COL.IElement;
END_VAR
END_METHOD

METHOD ELEMENTEQUALS : BOOL
VAR_INPUT
	ITFELEMENT : COL.IElement;
END_VAR
END_METHOD

METHOD ELEMENTHASHCODE : LINT
END_METHOD

METHOD PRVINSTINIT : COL.FBF.ERROR
VAR_INPUT
	ITFDATA : COL.FBF.IData;
END_VAR
END_METHOD

(* ---- HASHTABLEVALUEELEMENTDATA.pou ---- *)
FUNCTION_BLOCK HASHTABLEVALUEELEMENTDATA EXTENDS InstanceData
VAR_INPUT
	UDIALARMGROUPID : UDINT;
	UITEMPLATEALARMSOFFSET : UINT;
	UITEMPLATEALARMSLENGTH : UINT;
	UITEMPLATEEVENTSOFFSET : UINT;
	UITEMPLATEEVENTSLENGTH : UINT;
END_VAR
END_FUNCTION_BLOCK

(* ---- HASHTABLEVALUEELEMENTFACTORY.pou ---- *)
FUNCTION_BLOCK HASHTABLEVALUEELEMENTFACTORY EXTENDS FactoryBase
VAR
	PRVINSTCOUNT : CAA.COUNT;
	PRVINSTPOOLEXTENDSFACTOR : USINT;
	PRVINSTSIZE : CAA.SIZE;
END_VAR
END_FUNCTION_BLOCK

METHOD CREATE : IHashtableValueElement
VAR_INPUT
	UDIALARMGROUPID : UDINT;
	UITEMPLATEALARMSOFFSET : UINT;
	UITEMPLATEALARMSLENGTH : UINT;
	UITEMPLATEEVENTSOFFSET : UINT;
	UITEMPLATEEVENTSLENGTH : UINT;
END_VAR
VAR_OUTPUT
	EERROR : COL.FBF.ERROR;
END_VAR
END_METHOD

(* ---- HISTORICALALARMMOCK.pou ---- *)
FUNCTION_BLOCK HISTORICALALARMMOCK EXTENDS ProxyFbAlarmHistorical
VAR_INPUT
	M_BALARMSTORAGE : BYTE;
	M_DWROWIDFIRST : DWORD;
	M_DWROWIDLAST : DWORD;
	M_SVALUE : STRING;
	M_WSVALUE : WSTRING;
END_VAR
END_FUNCTION_BLOCK

METHOD SETVALUES
VAR_INPUT
	ISET : INT;
END_VAR
END_METHOD

(* ---- LISTELEMENT.pou ---- *)
FUNCTION_BLOCK LISTELEMENT EXTENDS InstanceBase
VAR
	_ALARMINST : Alarm;
	_USICOUNTLATCHVARIABLES : USINT;
	_ARRLATCHVARIABLES : ARRAY [0..255] OF ValueTypeBundle;
	_XISACTIVEALARM : BOOL;
	ALARM : POINTER TO Alarm;
	ISACTIVEALARM : BOOL;
	ISDEACTIVATEDPREV : BOOL;
END_VAR
END_FUNCTION_BLOCK

METHOD ELEMENTCOMPARETO : INT
VAR_INPUT
	ITFELEMENT : COL.IElement;
END_VAR
END_METHOD

METHOD ELEMENTEQUALS : BOOL
VAR_INPUT
	ITFELEMENT : COL.IElement;
END_VAR
END_METHOD

METHOD ELEMENTHASHCODE : LINT
END_METHOD

METHOD GETLATCHVARIABLES : BOOL
VAR_OUTPUT
	PALATCHVARIABLES : POINTER TO ARRAY [0..255] OF ValueTypeBundle;
	USICOUNTLATCHVARIABLES : USINT;
END_VAR
END_METHOD

METHOD SETLATCHVARIABLES : BOOL
VAR_INPUT
	PALARM : POINTER TO Alarm;
END_VAR
END_METHOD

METHOD PRVINSTINIT : COL.FBF.ERROR
VAR_INPUT
	ITFDATA : COL.FBF.IData;
END_VAR
END_METHOD

(* ---- LISTELEMENTDATA.pou ---- *)
FUNCTION_BLOCK LISTELEMENTDATA EXTENDS InstanceData
END_FUNCTION_BLOCK

(* ---- LISTELEMENTFACTORY.pou ---- *)
FUNCTION_BLOCK LISTELEMENTFACTORY EXTENDS FactoryBase
VAR
	PRVINSTCOUNT : CAA.COUNT;
	PRVINSTPOOLEXTENDSFACTOR : USINT;
	PRVINSTSIZE : CAA.SIZE;
END_VAR
END_FUNCTION_BLOCK

METHOD CREATE : IListElement
VAR_OUTPUT
	EERROR : COL.FBF.ERROR;
END_VAR
END_METHOD

(* ---- MESSAGECOMPARER.pou ---- *)
FUNCTION_BLOCK MESSAGECOMPARER EXTENDS TSLastComparer
VAR
	M_STRINGTYPE : __SYSTEM.TYPE_CLASS;
	M_IWHICHMESSAGE : INT;
	M_ICOUNTLATCHVARIABLES : INT;
	M_CBSMESSAGE1 : CharBufferString;
	M_CBSMESSAGE2 : CharBufferString;
	M_CBSMESSAGE1REPLACED : CharBufferString;
	M_CBSMESSAGE2REPLACED : CharBufferString;
	M_ABYBUFFERMESSAGE1REPLACED : ARRAY [0..(BUFFER_LENGTH - 1)] OF BYTE;
	M_ABYBUFFERMESSAGE2REPLACED : ARRAY [0..(BUFFER_LENGTH - 1)] OF BYTE;
	M_TIMESTAMPANDVALUESCONTAINER : TimestampAndValuesContainer;
	BUFFER_LENGTH : INT := (2 * (255 + 1));
END_VAR
END_FUNCTION_BLOCK

METHOD BEFORECOMPARE
VAR_INPUT
	STRINGTYPE : __SYSTEM.TYPE_CLASS;
	IWHICHMESSAGE : INT;
	ICOUNTLATCHVARIABLES : INT;
END_VAR
END_METHOD

METHOD COMPARE : INT
VAR_INPUT
	DIINDEXALARM1 : DINT;
	DIINDEXALARM2 : DINT;
END_VAR
END_METHOD

METHOD PRVGETALARMMESSAGE : CharBufferPtr
VAR_INPUT
	UDIALARMGROUPID : UDINT;
	UDIALARMID : UDINT;
	SDEVICENAME : STRING;
END_VAR
VAR_OUTPUT
	SALARMID : STRING;
END_VAR
END_METHOD

METHOD PRVREPLACEPLACEHOLDERS : BOOL
VAR_INPUT
	DIINDEXALARM : DINT;
	CBPMESSAGE : CharBufferPtr;
	RCBSMESSAGE : REFERENCE TO CharBufferString;
	RCBSMESSAGEREPLACED : REFERENCE TO CharBufferString;
END_VAR
END_METHOD

(* ---- ONLYDATEANDTIMEPLACEHOLDER.pou ---- *)
FUNCTION_BLOCK ONLYDATEANDTIMEPLACEHOLDER
VAR
	M_APLACEHOLDEROCCURRENCE : ARRAY [PLACEHOLDER_DATE..PLACEHOLDER_TIME] OF PlaceholderOccurrence;
	PLACEHOLDER_DATE : INT := 0;
	PLACEHOLDER_TIME : INT := 1;
END_VAR
END_FUNCTION_BLOCK

METHOD FB_INIT : BOOL
VAR_INPUT
	BINITRETAINS : BOOL;
	BINCOPYCODE : BOOL;
END_VAR
END_METHOD

METHOD ANALYZEPLACEHOLDERS
VAR_INPUT
	STRINGTYPE : __SYSTEM.TYPE_CLASS;
END_VAR
END_METHOD

METHOD GETCOUNTPLACEHOLDERS : SINT
END_METHOD

METHOD GETPLACEHOLDER : PlaceholderOccurrence
VAR_INPUT
	SIWHICHPLACEHOLDER : SINT;
END_VAR
END_METHOD

METHOD HASPLACEHOLDERREQUIRINGCYCLICALLYUPDATE : BOOL
END_METHOD

METHOD HASPLACEHOLDERS : BOOL
END_METHOD

METHOD ISOPTIMIZEDPLACEHOLDERREPLACEMENTSUPPORTED : BOOL
END_METHOD

(* ---- PRIORITYCOMPARER.pou ---- *)
FUNCTION_BLOCK PRIORITYCOMPARER EXTENDS TSLastComparer
END_FUNCTION_BLOCK

METHOD COMPARE : INT
VAR_INPUT
	DIINDEXALARM1 : DINT;
	DIINDEXALARM2 : DINT;
END_VAR
END_METHOD

(* ---- PROXY.pou ---- *)
FUNCTION_BLOCK PROXY
VAR
	M_XISINIT : BOOL;
	M_IRUNSTATUS : INT;
	M_ITFCOMMCHANNEL : IProxyCommChannel;
	M_ITEST : INT;
	M_ESTATE : ProxyEnumState;
	M_SDEVICENAME : STRING;
	M_LIBVERALMMAN : VERSION;
	M_LTSTARTTIMECHANNEL : LTIME;
	M_LTSTARTTIMERUN : LTIME;
	M_LTSTARTTIME : LTIME;
	M_ISTATE : INT;
	M_XALREADYDISP : BOOL;
	M_TTIMEOUT : TIME;
	M_IREQIDSENT : INT;
	M_IREQIDREC : INT;
	M_XWITHERRORS : BOOL;
	M_DWBASETIME : DWORD := (50 * 1000);
	M_DWACTALMTIME : DWORD := (200 * 1000);
	M_DWHISALMTIME : DWORD := (1000 * 1000);
	M_DWACKALMTIME : DWORD := (1000 * 1000);
	M_TGENTIMEOUT : TIME := DEFAULT_TIMEOUT;
	M_APROXYRUNTASKCALL : ARRAY [1..ProxyConstants.MAX_TASK] OF ProxyStructTaskCall;
	M_IRUNTASKCALLMAX : INT;
	M_APROXYPRERUNTASKCALL : ARRAY [1..ProxyConstants.MAX_TASK] OF ProxyStructTaskCall;
	M_IPRERUNTASKCALLMAX : INT;
	M_ITASKCALL : INT;
	M_SPROXYNAME : STRING;
	M_PSAPPNAME : POINTER TO STRING;
	M_CBSMESSAGE : CharBufferString;
	M_AWLOCALBUFFER : ARRAY [0..(LOCAL_TEXT_BUFFER_LENGTH / 2)] OF WORD;
	M_ARECORDS : ARRAY [0..(MAX_RECORDS - 1)] OF ProxyStructRecord;
	M_IRECINUSE : INT;
	M_SIHASSTORAGE : SINT := -1;
	M_DWROWIDFIRSTREMDB : DWORD := AlarmConstants.INVALID_ROWID;
	M_DWROWIDLASTREMDB : DWORD := AlarmConstants.INVALID_ROWID;
	M_DWROWIDLASTVALIDREAD : DWORD := AlarmConstants.INVALID_ROWID;
	M_DWROWIDLASTLOCDB : DWORD := AlarmConstants.INVALID_ROWID;
	M_IROWCOUNTTOREAD : INT;
	M_PAHISTALARMGROUPS : ARRAY [1..MAX_HIST_GROUPS] OF POINTER TO STRING;
	M_IHISTALARMGROUPSNUM : INT;
	M_IHISTRECORDID : INT := -1;
	M_XFIRSTHISTREADDONE : BOOL;
	M_XFIRSTHISTACTIVEREADDONE : BOOL;
	M_XDISP1DONE : BOOL;
	M_XDISP2DONE : BOOL;
	M_XDISP3DONE : BOOL;
	M_XDISP4DONE : BOOL;
	M_DIHISTACTIVEFIRSTENTRY : DINT;
	M_HISTACTIVEALMPENDINGQUEUE : ProxyFbHistActiveAlarmsQueue;
	M_HISTALMROWQUEUE : ProxyFbHistAlarmsRowQueue;
	M_HISTACTIVEALMROWQUEUE : ProxyFbHistAlarmsRowQueue;
	M_IHISTROWCOUNTREAD : INT;
	M_IHISTACTIVEROWCOUNTREAD : INT;
	M_TWRITEDBDURATIONTIME : TIME;
	M_IWRITEDBCNT : INT;
	M_DIWRITEDBCNTTOT : DINT;
	M_DISTORAGEROWSCOUNT : DINT;
	M_ISTORAGECLEAR : INT;
	M_ISTORAGECLEAROLD : INT := -1;
	M_IRECIXALMTOACK : INT;
	M_DIALMIXALMTOACK : DINT;
	M_LITIMELASTLOCDB : LINT;
	M_IVERSIONDB : INT;
	M_XCLIENTISREG : BOOL;
	M_HLOCKREADALM2 : RTS_IEC_HANDLE := RTS_INVALID_HANDLE;
	M_ICNTFORSTATISTICS : INT;
	M_DISTATHISTACTIVEALMSCNT : DINT;
	M_ISTATHISTROWALMSCNT : INT;
	M_ISTATHISTROWACTIVEALMSCNT : INT;
	_IRECORDID : INT;
	_DIALARMNUM : DINT;
	_ILATCHVARSNUM : INT;
	_IALARMCLASSNUM : INT;
	_XRAISEDMOREALARMSTHANSTORAGELIMITREPORTED : BOOL;
	STATE_IDLE : INT := 0;
	STATE_ANS_WAIT : INT := 10;
	RUN_START : INT := 0;
	RUN_RECORD : INT := 1;
	RUN_RECORD_HIST : INT := 2;
	RUN_PRERUN : INT := 3;
	RUN_CHECK_DATA : INT := 4;
	RUN_RUN : INT := 5;
	MAX_RECORDS : INT := 1;
	MAX_HIST_GROUPS : INT := 50;
	DEFAULT_NAME : STRING := '-Proxy-';
	DEFAULT_TIMEOUT : TIME := TIME#30s0ms;
	LOCAL_TEXT_BUFFER_LENGTH : INT := (1000 * 2);
	ACTIVEALARMSCOUNT : DINT;
	APPLICATION : POINTER TO STRING;
	HASSTORAGE : BOOL;
	HISTACTIVEALARMREAD : INT;
	HISTALARMREAD : INT;
	ISINITIALIZED : BOOL;
	ISRUNCYCLICOK : BOOL;
	LATCHVARSNUM : INT;
	MAXHISTROWSTOREAD : INT;
	PROXYTASKCALL : ARRAY [1..ProxyConstants.MAX_TASK] OF ProxyStructTaskCall;
	PROXYTASKCALLSIZE : INT;
	RECORDID : INT;
	RECORDIDHISTORICAL : INT;
	ROWIDFIRST : DWORD;
	ROWIDLAST : DWORD;
	ROWIDLASTREAD : DWORD;
	TOTALARMNUM : DINT;
	TOTCLASSNUM : INT;
END_VAR
END_FUNCTION_BLOCK

METHOD FB_EXIT : BOOL
VAR_INPUT
	BINCOPYCODE : BOOL;
END_VAR
END_METHOD

METHOD FB_INIT : BOOL
VAR_INPUT
	BINITRETAINS : BOOL;
	BINCOPYCODE : BOOL;
END_VAR
END_METHOD

METHOD CYCLICCALL : BOOL
END_METHOD

METHOD GETACTIVEALARMS : INT
VAR_INPUT
	SNAME : STRING;
	FILTERCRITERIA : REFERENCE TO VisuFbAlarmFilterCriteria;
	ITFALARMDATABLOCK : IAlarmDataBlockBaseDINT;
END_VAR
VAR_IN_OUT
	DISTUBPROG : DINT;
END_VAR
END_METHOD

METHOD GETACTIVEALARMS2
VAR_INPUT
	FILTERCRITERIA : REFERENCE TO VisuFbAlarmFilterCriteria;
	PAITFALARMS : POINTER TO ARRAY [0..10] OF IAlarm;
	DIARRSIZE : DINT;
END_VAR
VAR_OUTPUT
	DICOUNT : DINT;
END_VAR
END_METHOD

METHOD GETALARMCLASSDESC
VAR_INPUT
	UDIID : UDINT;
END_VAR
VAR_OUTPUT
	SDESC : ProxyStructAlarmClassDesc;
END_VAR
END_METHOD

METHOD GETALARMCLASSDESCBYNAME
VAR_INPUT
	SCLASSNAME : STRING;
END_VAR
VAR_OUTPUT
	SDESC : ProxyStructAlarmClassDesc;
END_VAR
END_METHOD

METHOD GETALARMDESC
VAR_INPUT
	UDIALMID : UDINT;
	UDIGRPID : UDINT;
END_VAR
VAR_OUTPUT
	SDESC : ProxyStructAlarmDesc;
END_VAR
END_METHOD

METHOD GETALARMDISPLAYOPTIONS
VAR_INPUT
	ITFALARMMETAOBJECTSTUB5 : IAlarmMetaObjectStub5;
	REFDISPLAYOPTIONS : REFERENCE TO DisplayOptions;
END_VAR
VAR_OUTPUT
	XVALID : BOOL;
	SCLASSREMAP : STRING;
END_VAR
END_METHOD

METHOD GETALARMGROUPDESC
VAR_INPUT
	UDIID : UDINT;
END_VAR
VAR_OUTPUT
	SDESC : ProxyStructAlarmGroupDesc;
END_VAR
END_METHOD

METHOD GETALARMGROUPDESCBYNAME
VAR_INPUT
	SGRPNAME : STRING;
END_VAR
VAR_OUTPUT
	SDESC : ProxyStructAlarmGroupDesc;
END_VAR
END_METHOD

METHOD GETALARMMESSAGE
VAR_INPUT
	ITFALARMMETAOBJECTSTUB5 : IAlarmMetaObjectStub5;
	IWHICHMESSAGE : INT;
	REFCHARBUFFERSTRING : REFERENCE TO CharBufferString;
	STRINGTYPE : __SYSTEM.TYPE_CLASS;
END_VAR
END_METHOD

METHOD GETALARMMESSAGE2 : Stu.CharBufferPtr
VAR_INPUT
	STEXTLISTNAME : STRING;
	STEXTLISTINDEX : STRING;
	IWHICHMESSAGE : INT;
	STRINGTYPE : __SYSTEM.TYPE_CLASS;
END_VAR
END_METHOD

METHOD GETPROXYNAME : POINTER TO STRING
END_METHOD

METHOD GETTOTALALARMSCOUNT : DINT
END_METHOD

METHOD INITIALIZE : BOOL
VAR_INPUT
	PPARAM : POINTER TO ProxyStructInitialize;
	ITEST : INT;
END_VAR
END_METHOD

METHOD REGISTERUSERCLIENT
END_METHOD

METHOD SETALARMSTOACK
VAR_INPUT
	ITFALARMMETAOBJECTSTUB : IAlarmMetaObjectStub5;
END_VAR
END_METHOD

METHOD SETINITIALDATAFROMDB
VAR_INPUT
	ROW : REFERENCE TO AlarmStorageRow;
	XFIRST : BOOL;
	IVERSION : INT;
END_VAR
END_METHOD

METHOD SETPARAMS
VAR_INPUT
	PPARAM : POINTER TO ProxyStructParam;
END_VAR
END_METHOD

METHOD COMMUNICATIONFINISHED
VAR_INPUT
	IREQUESTID : INT;
	XWITHERRORS : BOOL;
END_VAR
END_METHOD

METHOD PROXYMANAGERLOG
VAR_INPUT
	SVAL1 : STRING(255);
	SVAL2 : STRING(255);
	SVAL3 : STRING(255);
	UDISEV : UDINT;
END_VAR
END_METHOD

METHOD SETACTIVEALARMSCOUNT
VAR_INPUT
	DICOUNT : DINT;
END_VAR
END_METHOD

METHOD SETALARMMANAGERLIBVERSION
VAR_INPUT
	LIBVER : VERSION;
END_VAR
END_METHOD

METHOD SETDEVICENAME
VAR_INPUT
	SNAME : STRING;
END_VAR
END_METHOD

METHOD SETHASSTORAGE
VAR_INPUT
	XVALUE : BOOL;
END_VAR
END_METHOD

METHOD SETHISTACTIVEALARMSREAD
VAR_INPUT
	ICOUNT : INT;
END_VAR
END_METHOD

METHOD SETHISTALARMSREAD
VAR_INPUT
	DWROWIDLAST : DWORD;
	ICOUNT : INT;
	DISTORAGEROWSCOUNT : DINT;
	ISTORAGECLEAR : INT;
END_VAR
END_METHOD

METHOD SETLATCHVARSCOUNT
VAR_INPUT
	ICOUNT : INT;
END_VAR
END_METHOD

METHOD SETRECORDID
VAR_INPUT
	IVALUE : INT;
END_VAR
END_METHOD

METHOD SETROWIDS
VAR_INPUT
	DWROWIDFIRST : DWORD;
	DWROWIDLAST : DWORD;
END_VAR
END_METHOD

METHOD SETTOTALALARMSCOUNT
VAR_INPUT
	DICOUNT : DINT;
END_VAR
END_METHOD

METHOD SETTOTALCLASSESCOUNT
VAR_INPUT
	ICOUNT : INT;
END_VAR
END_METHOD

METHOD GETALARMGROUP : STRING
VAR_INPUT
	IWHICHALARMGROUP : INT;
END_VAR
END_METHOD

METHOD GETALARMGROUPSNUM : INT
END_METHOD

METHOD GETAPPLICATION : STRING
END_METHOD

METHOD GETCOUNTALARMSTOACKNOWLEDGE : INT
END_METHOD

METHOD GETNEXTALARMTOACKNOWLEDGE : BOOL
VAR_INPUT
	XFISRTENTRY : BOOL;
END_VAR
VAR_OUTPUT
	ALARMTOACKNOWLEDGE : AlarmToAcknowledge;
END_VAR
END_METHOD

METHOD GETPROXYACTIVEALARMOBJECT : IProxyAlarmObject
VAR_INPUT
	DIOBJNUM : DINT;
END_VAR
END_METHOD

METHOD GETPROXYALARMCLASSDESCRIPTIONOBJECT : POINTER TO ProxyStructAlarmClass
VAR_INPUT
	IOBJNUM : INT;
END_VAR
END_METHOD

METHOD GETPROXYALARMDESCRIPTIONOBJECT : POINTER TO ProxyStructAlarm
VAR_INPUT
	IOBJNUM : INT;
END_VAR
END_METHOD

METHOD GETPROXYALARMGROUPDESCRIPTIONOBJECT : POINTER TO ProxyStructAlarmGroup
VAR_INPUT
	IOBJNUM : INT;
END_VAR
END_METHOD

METHOD GETPROXYHISTORICALALARMOBJECT : POINTER TO ProxyFbAlarmHistorical
VAR_INPUT
	XACTIVE : BOOL;
	IOBJNUM : INT;
END_VAR
END_METHOD

METHOD GETRECORDID : INT
END_METHOD

METHOD GETRECORDIDHISTORICAL : INT
END_METHOD

METHOD GETROWIDHISTORICALACTIVEALARMS
VAR_INPUT
	XFIRSTCALL : BOOL;
END_VAR
VAR_OUTPUT
	DWROWID : DWORD;
	LITS : LINT;
END_VAR
END_METHOD

METHOD GETROWTOREAD
VAR_OUTPUT
	DWROWIDLAST : DWORD;
	IROWCOUNT : INT;
END_VAR
END_METHOD

METHOD PRVCHECKALARMCLASS
VAR_INPUT
	PRECORDDATA : POINTER TO ProxyStructRecord;
END_VAR
END_METHOD

METHOD PRVCHECKALARMGROUP
VAR_INPUT
	PRECORDDATA : POINTER TO ProxyStructRecord;
END_VAR
END_METHOD

METHOD PRVGETALARMCLASSDESC : POINTER TO ProxyStructAlarmClass
VAR_INPUT
	PRECORDDATA : POINTER TO ProxyStructRecord;
	UICLASSID : UDINT;
END_VAR
END_METHOD

METHOD PRVGETALARMCLASSDESCBYNAME : POINTER TO ProxyStructAlarmClass
VAR_INPUT
	PRECORDDATA : POINTER TO ProxyStructRecord;
	SNAME : STRING;
END_VAR
END_METHOD

METHOD PRVGETALARMCONTAINER : POINTER TO AlarmContainer
VAR_INPUT
	DIOBJNUM : DINT;
	PSTRURECORD : POINTER TO ProxyStructRecord;
END_VAR
END_METHOD

METHOD PRVGETALARMDESC : POINTER TO ProxyStructAlarm
VAR_INPUT
	PRECORDDATA : POINTER TO ProxyStructRecord;
	UIALARMID : ALARM_ID;
	UDIGROUPID : UDINT;
END_VAR
END_METHOD

METHOD PRVGETALARMDESC2 : POINTER TO ProxyStructAlarm
VAR_INPUT
	PRECORDDATA : POINTER TO ProxyStructRecord;
	UDIALARMINTERNALID : UDINT;
	UDIGROUPID : UDINT;
END_VAR
END_METHOD

METHOD PRVGETALARMGROUPDESC : POINTER TO ProxyStructAlarmGroup
VAR_INPUT
	PSTRURECORD : POINTER TO ProxyStructRecord;
	UDIID : UDINT;
END_VAR
END_METHOD

METHOD PRVGETLOCK : RTS_IEC_HANDLE
VAR_INPUT
	ITASKID : INT;
END_VAR
END_METHOD

METHOD PRVGETPROXYACTIVEALARMOBJECT : IProxyAlarmObject
VAR_INPUT
	DIOBJNUM : DINT;
	PSTRURECORD : POINTER TO ProxyStructRecord;
END_VAR
END_METHOD

METHOD PRVGETRECORDDATA : POINTER TO ProxyStructRecord
VAR_INPUT
	IINDEX : INT;
END_VAR
END_METHOD

METHOD PRVPREPAREFORRESTART
END_METHOD

METHOD GETALARMCLASSESDESCRIPTION
VAR_INPUT
	PCLDESC : POINTER TO ARRAY [0..0] OF ProxyStructMonitorAlarmClassDesc;
	ISIZE : INT;
END_VAR
VAR_OUTPUT
	ICLCNT : INT;
END_VAR
END_METHOD

METHOD GETALARMGROUPSDESCRIPTION
VAR_INPUT
	PGRPDESC : POINTER TO ARRAY [0..0] OF ProxyStructMonitorAlarmGroupDesc;
	ISIZE : INT;
END_VAR
VAR_OUTPUT
	IGRPCNT : INT;
END_VAR
END_METHOD

METHOD GETALARMSDESCRIPTION
VAR_INPUT
	PALMDESC : POINTER TO ARRAY [0..0] OF ProxyStructMonitorAlarmDesc;
	DISIZE : DINT;
END_VAR
VAR_OUTPUT
	DIALMCNT : DINT;
END_VAR
END_METHOD

METHOD GETSTATISTICS : ProxyStructMonitor
VAR_INPUT
	IRECORD : INT;
END_VAR
END_METHOD

METHOD GETSTATISTICSSINGLEREQ : ProxyStructMonitorRequest
VAR_INPUT
	ITASKID : INT;
END_VAR
END_METHOD

METHOD PRVREADHISTALARMSPREELAB : SINT
VAR_INPUT
	IREQID : INT;
END_VAR
END_METHOD

METHOD PRVALARMOBJECTALLOC
VAR_INPUT
	PSTRURECORD : POINTER TO ProxyStructRecord;
END_VAR
END_METHOD

METHOD PRVALARMOBJECTFREE
VAR_INPUT
	PSTRURECORD : POINTER TO ProxyStructRecord;
END_VAR
END_METHOD

METHOD PRVALARMOBJECTSTUBSALLOC
VAR_INPUT
	PSTRURECORD : POINTER TO ProxyStructRecord;
END_VAR
END_METHOD

METHOD PRVALARMOBJECTSTUBSFREE
VAR_INPUT
	PSTRURECORD : POINTER TO ProxyStructRecord;
END_VAR
END_METHOD

METHOD PRVSTRUCTALARMCLASSDESCRIPTIONALLOC
VAR_INPUT
	PSTRURECORD : POINTER TO ProxyStructRecord;
END_VAR
END_METHOD

METHOD PRVSTRUCTALARMCLASSDESCRIPTIONFREE
VAR_INPUT
	PSTRURECORD : POINTER TO ProxyStructRecord;
END_VAR
END_METHOD

METHOD PRVSTRUCTALARMDESCRIPTIONALLOC
VAR_INPUT
	PSTRURECORD : POINTER TO ProxyStructRecord;
END_VAR
END_METHOD

METHOD PRVSTRUCTALARMDESCRIPTIONFREE
VAR_INPUT
	PSTRURECORD : POINTER TO ProxyStructRecord;
END_VAR
END_METHOD

METHOD PRVSTRUCTALARMGROUPDESCRIPTIONALLOC
VAR_INPUT
	PSTRURECORD : POINTER TO ProxyStructRecord;
END_VAR
END_METHOD

METHOD PRVSTRUCTALARMGROUPDESCRIPTIONFREE
VAR_INPUT
	PSTRURECORD : POINTER TO ProxyStructRecord;
END_VAR
END_METHOD

METHOD PRVGETENTRYTASKCALLTABLE : POINTER TO ProxyStructTaskCall
VAR_INPUT
	ITASKID : INT;
	ITABLE : INT;
END_VAR
END_METHOD

METHOD PRVPREPAREPRERUNTASKCALLTABLE
END_METHOD

METHOD PRVPREPARERUNTASKCALLTABLE
END_METHOD

(* ---- PROXYDATASOURCECHANNEL.pou ---- *)
FUNCTION_BLOCK PROXYDATASOURCECHANNEL
VAR
	M_ITFDATASOURCESMGR : IDatasources.IDatasourcesMgr;
	M_PSDSNAME : POINTER TO STRING;
	M_DIALARMNUM : DINT;
	M_IALARMCLASSNUM : INT;
	M_ILATCHVARSNUM : INT;
	M_ITFDATASOURCE : IDatasources.IDatasource2;
	M_IMAXALMGROUPS : INT;
	M_PSALMSTATETRANSCOUNTER : POINTER TO STRING;
	M_PALMSTATETRANSCOUNTER : __XWORD;
	M_TYPEALMSTATETRANSCOUNTER : TypeClass;
	M_XALMSTATETRANSCOUNTERISREG : BOOL;
	M_LIOLDSTATETRANSCOUNTERVALUE : LINT := -1;
	M_PSALMSTORAGECOUNTER : POINTER TO STRING;
	M_PALMSTORAGECOUNTER : __XWORD;
	M_TYPEALMSTORAGECOUNTER : TypeClass;
	M_XALMSTORAGECOUNTERISREG : BOOL;
	M_LIOLDSTORAGECOUNTERVALUE : LINT := -1;
	M_LIOLDSTORAGECOUNTERVALUE2 : LINT := -1;
	M_REQUESTBUILDERSETALMRECORD : RequestBuilderSetAlmRecord;
	M_REQUESTBUILDERRESALMRECORD : RequestBuilderResetAlmRecord;
	M_REQUESTBUILDERREADACTIVEALARMS : RequestBuilderReadActiveAlarms;
	M_REQUESTBUILDERGETALMCONFIG : RequestBuilderGetAlmConfig;
	M_REQUESTBUILDERGETALMCLASSCONFIG : RequestBuilderGetAlmClassConfig;
	M_REQUESTBUILDERACKALARMS : RequestBuilderAckAlarms;
	M_REQUESTBUILDERGETHISTORICALALMCONFIG : RequestBuilderGetHistoricalAlmConfig;
	M_REQUESTBUILDERREADHISTORICALALARMS : RequestBuilderReadHistoricalAlarms;
	M_REQUESTBUILDERREADHISTORICALACTIVEALARMS : RequestBuilderReadHistoricalActiveAlarms;
	M_REQUESTBUILDERCHANNELTEST : RequestBuilderChannelTest;
	M_REQUESTBUILDERCHANNELTEST2 : RequestBuilderChannelTest2;
	M_ITFPROXYCONSUMER : IProxyConsumer;
	M_ITFPROXYPROVIDER : IProxyProvider;
	M_ICURRREQUESTID : INT;
	M_ICOUNTTEST : INT;
	M_IERRORFROMDEV : INT;
	M_IHISTROWCOUNTREAD : INT;
	M_IHISTACTIVEROWCOUNTREAD : INT;
	M_IROWCOUNTREAD : INT;
	M_PFBREQUESTCALLED : POINTER TO RequestBuilderBase;
	M_XFIRSTCALL : BOOL := TRUE;
	M_LTLASTREADACTALM : LTIME;
	M_LTLASTREADHISTALM : LTIME;
	M_LTLASTREADHISTACTALM : LTIME;
	_SDEVICENAME : STRING;
	_ILATCHVARSNUM : INT;
	_IRECORDID : INT;
	_XHASSTORAGE : BOOL;
	_DWROWIDFIRST : DWORD;
	_DWROWIDLAST : DWORD;
	ALMSTATETRANSCOUNTERREGISTERED : BOOL;
	ALMSTORAGECOUNTERREGISTERED : BOOL;
	DEVICENAME : STRING;
	ERRORFROMDEVICE : INT;
	HASSTORAGE : BOOL;
	LATCHVARSNUM : INT;
	RECORDID : INT;
	ROWIDFIRST : DWORD;
	ROWIDLAST : DWORD;
	TESTVARIABLEVALUE : INT;
	TOTALARMNUM : DINT;
	TOTCLASSNUM : INT;
END_VAR
END_FUNCTION_BLOCK

METHOD SETPARAMS
VAR_INPUT
	PPARAM : POINTER TO ProxyStructDSChannelParam;
END_VAR
END_METHOD

METHOD GETCOUNTALARMSTOACKNOWLEDGE : INT
END_METHOD

METHOD GETNEXTALARMTOACKNOWLEDGE : BOOL
VAR_INPUT
	XFISRTENTRY : BOOL;
END_VAR
VAR_OUTPUT
	ALARMTOACKNOWLEDGE : AlarmToAcknowledge;
END_VAR
END_METHOD

METHOD GETPROXYALARMCLASSDESCRIPTIONOBJECT : POINTER TO ProxyStructAlarmClass
VAR_INPUT
	IOBJNUM : INT;
END_VAR
END_METHOD

METHOD GETPROXYALARMDESCRIPTIONOBJECT : POINTER TO ProxyStructAlarm
VAR_INPUT
	IOBJNUM : INT;
END_VAR
END_METHOD

METHOD GETPROXYALARMGROUPDESCRIPTIONOBJECT : POINTER TO ProxyStructAlarmGroup
VAR_INPUT
	IOBJNUM : INT;
END_VAR
END_METHOD

METHOD SETALARMMANAGERLIBVERSION
VAR_INPUT
	LIBVER : VERSION;
END_VAR
END_METHOD

METHOD SETALARMSCOUNT
VAR_INPUT
	DIVALUE : DINT;
END_VAR
END_METHOD

METHOD SETCLASSESCOUNT
VAR_INPUT
	IVALUE : INT;
END_VAR
END_METHOD

METHOD SETRECORDID
VAR_INPUT
	IVALUE : INT;
END_VAR
END_METHOD

METHOD GETALARMGROUP : STRING
VAR_INPUT
	IWHICHALARMGROUP : INT;
END_VAR
END_METHOD

METHOD GETALARMGROUPSNUM : INT
END_METHOD

METHOD SETVALUE
VAR_INPUT
	IVALUE : INT;
END_VAR
END_METHOD

METHOD GETVALUE : INT
END_METHOD

METHOD SETHASSTORAGE
VAR_INPUT
	XVALUE : BOOL;
END_VAR
END_METHOD

METHOD SETHISTACTIVEALARMSREAD
VAR_INPUT
	ICOUNT : INT;
END_VAR
END_METHOD

METHOD SETHISTALARMSREAD
VAR_INPUT
	DWROWIDLAST : DWORD;
	ICOUNT : INT;
	DISTORAGEROWSCOUNT : DINT;
	ISTORAGECLEAR : INT;
END_VAR
END_METHOD

METHOD SETROWIDS
VAR_INPUT
	DWROWIDFIRST : DWORD;
	DWROWIDLAST : DWORD;
END_VAR
END_METHOD

METHOD GETPROXYHISTORICALALARMOBJECT : POINTER TO ProxyFbAlarmHistorical
VAR_INPUT
	XACTIVE : BOOL;
	IOBJNUM : INT;
END_VAR
END_METHOD

METHOD GETRECORDIDHISTORICAL : INT
END_METHOD

METHOD GETROWIDHISTORICALACTIVEALARMS
VAR_INPUT
	XFIRSTCALL : BOOL;
END_VAR
VAR_OUTPUT
	DWROWID : DWORD;
	LITS : LINT;
END_VAR
END_METHOD

METHOD GETROWTOREAD
VAR_OUTPUT
	DWROWIDLAST : DWORD;
	IROWCOUNT : INT;
END_VAR
END_METHOD

METHOD ADDERROR
VAR_INPUT
	ITASKID : INT;
	UDIERROR : UDINT;
	SMSG : STRING;
END_VAR
END_METHOD

METHOD CLEANSTATISTICS : BOOL
VAR_INPUT
	ITASKID : INT;
END_VAR
END_METHOD

METHOD CYCLICCALL
END_METHOD

METHOD EXECUTEREQUEST : UDINT
VAR_INPUT
	ITASKID : INT;
	XLOCK : BOOL;
	HLOCK : RTS_IEC_HANDLE;
END_VAR
END_METHOD

METHOD GETALARMMESSAGETEXT : BOOL
VAR_INPUT
	ITFALARMMETAOBJECTSTUB5 : IAlarmMetaObjectStub5;
	IWHICHMESSAGE : INT;
	STRINGTYPE : __SYSTEM.TYPE_CLASS;
END_VAR
VAR_OUTPUT
	CBPMESSAGE : CharBufferPtr;
END_VAR
END_METHOD

METHOD GETALARMMESSAGETEXT2 : BOOL
VAR_INPUT
	STEXTLISTNAME : STRING;
	STEXTLISTINDEX : STRING;
	IWHICHMESSAGE : INT;
	STRINGTYPE : __SYSTEM.TYPE_CLASS;
END_VAR
VAR_OUTPUT
	CBPMESSAGE : CharBufferPtr;
END_VAR
END_METHOD

METHOD GETSTATISTICSSINGLEREQ : ProxyStructMonitorRequest
VAR_INPUT
	ITASKID : INT;
END_VAR
END_METHOD

METHOD INITIALIZE
VAR_INPUT
	ITFPROXYCONSUMER : IProxyConsumer;
	ITFPROXYPROVIDER : IProxyProvider;
	IMAXALMGROUPS : INT;
END_VAR
END_METHOD

METHOD ISCHANNELAVAILABLE : BOOL
END_METHOD

METHOD ISREQUESTEXECUTABLE : BOOL
VAR_INPUT
	ITASKID : INT;
	XTRYTOFORCE : BOOL;
END_VAR
END_METHOD

METHOD RESTART
END_METHOD

METHOD SETACTIVEALARMSCOUNT
VAR_INPUT
	DICOUNT : DINT;
END_VAR
END_METHOD

METHOD GETPROXYACTIVEALARMOBJECT : IProxyAlarmObject
VAR_INPUT
	DIOBJNUM : DINT;
END_VAR
END_METHOD

METHOD ERRORADDED
VAR_INPUT
	UDIERROR : UDINT;
	SMSG : STRING;
	STASKNAME : STRING;
END_VAR
END_METHOD

METHOD REQUESTCLOSED
VAR_INPUT
	IREQUESTID : INT;
END_VAR
END_METHOD

METHOD SETERRORFROMDEVICE
VAR_INPUT
	IERROR : INT;
END_VAR
END_METHOD

METHOD GETAPPLICATION : STRING
END_METHOD

METHOD GETDEVICENAME : STRING
END_METHOD

METHOD GETRECORDID : INT
END_METHOD

METHOD PRVGETALARMMESSAGETEXT
VAR_INPUT
	STEXTLISTNAME : STRING;
	STEXTLISTINDEX : STRING;
	IWHICHMESSAGE : INT;
	STRINGTYPE : __SYSTEM.TYPE_CLASS;
END_VAR
VAR_OUTPUT
	CBPMESSAGE : CharBufferPtr;
END_VAR
END_METHOD

METHOD PRVGETREQUESTBUILDERFB : POINTER TO RequestBuilderBase
VAR_INPUT
	ITASKID : INT;
END_VAR
END_METHOD

(* ---- PROXYFBALARMHISTORICAL.pou ---- *)
FUNCTION_BLOCK PROXYFBALARMHISTORICAL
VAR_INPUT
	M_DIHASTOREGISTERED : DINT;
	M_LATCHSTRINGS : ARRAY [1..MAX_LATCH_VARS] OF WSTRING;
	M_ROW : AlarmStorageRow;
END_VAR
VAR
	ALATCHVARIABLES : ARRAY [1..MAX_LATCH_VARS] OF LatchVariable;
	ALARMFB : Alarm;
END_VAR
END_FUNCTION_BLOCK

METHOD FB_INIT : BOOL
VAR_INPUT
	BINITRETAINS : BOOL;
	BINCOPYCODE : BOOL;
END_VAR
END_METHOD

(* ---- PROXYFBALARMMETAOBJECTSTUB.pou ---- *)
FUNCTION_BLOCK PROXYFBALARMMETAOBJECTSTUB
VAR_INPUT
	M_USILATCHVARSAVAIL : USINT;
END_VAR
VAR
	M_ALATCHVARIABLES : ARRAY [0..(MAX_LATCH_VARS - 1)] OF ValueTypeBundle;
	M_USICOUNTLATCHVARIABLES : USINT;
	M_UIID : ALARM_ID;
	M_UDIALARMGROUPINTERNALID : UDINT;
	M_LITIMESTAMPACKNOWLEDGE : AlarmManager_Interfaces.Timestamp;
	M_LITIMESTAMPACTIVE : AlarmManager_Interfaces.Timestamp;
	M_LITIMESTAMPINACTIVE : AlarmManager_Interfaces.Timestamp;
	M_LITIMESTAMPLAST : AlarmManager_Interfaces.Timestamp;
	M_IOFFSETACKNOWLEDGE : INT := -1;
	M_IOFFSETACTIVE : INT := -1;
	M_IOFFSETINACTIVE : INT := -1;
	M_IOFFSETLAST : INT := -1;
	M_ISTATE : INT;
	M_SALARMGROUP : STRING;
	M_STESTLISTNAME : STRING;
	M_SALARMCLASS : STRING;
	M_UDIALARMCLASSINTERNALID : UDINT;
	M_BYPRIORITY : BYTE;
	M_SALARMID : STRING;
	M_SPROXYNAME : STRING;
	M_CURRENTVALUE : ValueTypeBundle;
	M_TRIGGERVALUE : ValueTypeBundle;
	ALARMCLASSINTERNALID : UDINT;
	ALARMGROUPINTERNALID : UDINT;
	ALARMINTERNALID : UDINT;
	OFFSETACKNOWLEDGE : INT;
	OFFSETACTIVE : INT;
	OFFSETINACTIVE : INT;
	OFFSETLAST : INT;
	PROXYNAME : STRING;
END_VAR
END_FUNCTION_BLOCK

METHOD FB_EXIT : BOOL
VAR_INPUT
	BINCOPYCODE : BOOL;
END_VAR
END_METHOD

METHOD GETCHECKSUM : UDINT
END_METHOD

METHOD GETCURRENTVALUE : AlarmManagerInternal_Interfaces.ITypedValue
END_METHOD

METHOD SETACKNOWLEDGE
VAR_INPUT
	BACKNOWLEDGEMULTIPLE : BOOL;
END_VAR
END_METHOD

METHOD SWAPVALUES
END_METHOD

METHOD GETACKNOWLEDGE : BOOL
END_METHOD

METHOD GETACKNOWLEDGEMULTIPLE : BOOL
END_METHOD

METHOD GETALARMCLASS : STRING
END_METHOD

METHOD GETPRIORITY : BYTE
END_METHOD

METHOD GETSTRINGID : STRING
END_METHOD

METHOD GETTESTLISTNAME : STRING
END_METHOD

METHOD RESETACKNOWLEDGE
END_METHOD

METHOD SETALARMCLASS
VAR_INPUT
	SALARMCLASS : STRING;
END_VAR
END_METHOD

METHOD SETCURRENTVALUE
VAR_INPUT
	ITFTYPEDVALUECURRENT : AlarmManager_Interfaces.ITypedValue;
END_VAR
END_METHOD

METHOD SETPRIORITY
VAR_INPUT
	BYPRIORITY : BYTE;
END_VAR
END_METHOD

METHOD SETSTRINGID
VAR_INPUT
	SID : STRING;
END_VAR
END_METHOD

METHOD SETTESTLISTNAME
VAR_INPUT
	STESTLISTNAME : STRING;
END_VAR
END_METHOD

METHOD SETACKNOWLEDGE2
VAR_INPUT
	BACKNOWLEDGEMULTIPLE : BOOL;
END_VAR
END_METHOD

METHOD GETCOUNTLATCHVARIABLES : USINT
END_METHOD

METHOD GETLATCHVARVALUE : ITypedValue2
VAR_INPUT
	IWHICHLATCHVAR : INT;
END_VAR
END_METHOD

METHOD SETLATCHVARVALUE
VAR_INPUT
	IWHICHLATCHVAR : INT;
	ITFTYPEDVALUELATCHVAR : ITypedValue;
END_VAR
END_METHOD

METHOD SETCOUNTLATCHVARIABLES
VAR_INPUT
	USICOUNT : USINT;
END_VAR
END_METHOD

METHOD GETALARMGROUP : STRING
END_METHOD

METHOD GETID : AlarmManager_Interfaces.ALARM_ID
END_METHOD

METHOD GETLATCHVAR1VALUE : AlarmManager_Interfaces.ITypedValue
END_METHOD

METHOD GETLATCHVAR2VALUE : AlarmManager_Interfaces.ITypedValue
END_METHOD

METHOD GETSTATE : INT
END_METHOD

METHOD GETTIMESTAMPACKNOWLEDGE : AlarmManager_Interfaces.Timestamp
END_METHOD

METHOD GETTIMESTAMPACTIVE : AlarmManager_Interfaces.Timestamp
END_METHOD

METHOD GETTIMESTAMPINACTIVE : AlarmManager_Interfaces.Timestamp
END_METHOD

METHOD GETTIMESTAMPLAST : AlarmManager_Interfaces.Timestamp
END_METHOD

METHOD GETTRIGGERVALUE : AlarmManager_Interfaces.ITypedValue
END_METHOD

METHOD SETALARMGROUP
VAR_INPUT
	SALARMGROUP : STRING;
END_VAR
END_METHOD

METHOD SETID
VAR_INPUT
	UIID : AlarmManager_Interfaces.ALARM_ID;
END_VAR
END_METHOD

METHOD SETLATCHVAR1VALUE
VAR_INPUT
	ITFTYPEDVALUELATCHVAR1 : AlarmManager_Interfaces.ITypedValue;
END_VAR
END_METHOD

METHOD SETLATCHVAR2VALUE
VAR_INPUT
	ITFTYPEDVALUELATCHVAR2 : AlarmManager_Interfaces.ITypedValue;
END_VAR
END_METHOD

METHOD SETSTATE
VAR_INPUT
	ISTATE : INT;
END_VAR
END_METHOD

METHOD SETTIMESTAMPACKNOWLEDGE
VAR_INPUT
	LITIMESTAMPACKNOWLEDGE : AlarmManager_Interfaces.Timestamp;
END_VAR
END_METHOD

METHOD SETTIMESTAMPACTIVE
VAR_INPUT
	LITIMESTAMPACTIVE : AlarmManager_Interfaces.Timestamp;
END_VAR
END_METHOD

METHOD SETTIMESTAMPINACTIVE
VAR_INPUT
	LITIMESTAMPINACTIVE : AlarmManager_Interfaces.Timestamp;
END_VAR
END_METHOD

METHOD SETTIMESTAMPLAST
VAR_INPUT
	LITIMESTAMPLAST : AlarmManager_Interfaces.Timestamp;
END_VAR
END_METHOD

METHOD SETTRIGGERVALUE
VAR_INPUT
	ITFTYPEDVALUETRIGGER : AlarmManager_Interfaces.ITypedValue;
END_VAR
END_METHOD

(* ---- PROXYFBHISTACTIVEALARMSQUEUE.pou ---- *)
FUNCTION_BLOCK PROXYFBHISTACTIVEALARMSQUEUE
VAR
	M_PAALARM : POINTER TO ARRAY [0..10] OF POINTER TO ProxyStructHistoricalAlarmActive;
	M_DISZQUEUE : DINT;
	M_DISCANPOS : DINT;
	M_DICNTMAX : DINT;
	M_DICNT : DINT;
	M_DICNTAUX : DINT;
	SIZE_HIST_ACTIVE_ALARMS : INT := 50;
	EFFECTIVEREAD : DINT;
	QUEUESIZE : DINT;
END_VAR
END_FUNCTION_BLOCK

METHOD FB_EXIT : BOOL
VAR_INPUT
	BINCOPYCODE : BOOL;
END_VAR
END_METHOD

METHOD GETACTIVECOUNT : DINT
END_METHOD

METHOD GETAVAILABLEENTRIES : DINT
END_METHOD

METHOD GETLASTSTATE : AlarmState
VAR_INPUT
	DWROWID : DWORD;
END_VAR
END_METHOD

METHOD GETROWIDACTIVE
VAR_INPUT
	XFIRSTCALL : BOOL;
END_VAR
VAR_OUTPUT
	DWROWID : DWORD;
	LITS : LINT;
END_VAR
END_METHOD

METHOD GETROWIDLOCAL : DWORD
VAR_INPUT
	DWROWID : DWORD;
END_VAR
END_METHOD

METHOD INITIALIZE
END_METHOD

METHOD INSERT
VAR_INPUT
	SALM : ProxyStructHistoricalAlarmActive;
END_VAR
END_METHOD

METHOD ISPRESENTROWIDREMOTE : BOOL
VAR_INPUT
	DWROWID : DWORD;
END_VAR
END_METHOD

METHOD REMOVE
VAR_INPUT
	DWROWID : DWORD;
END_VAR
END_METHOD

METHOD SETLASTSTATE
VAR_INPUT
	DWROWID : DWORD;
	ESTATE : AlarmState;
END_VAR
END_METHOD

METHOD PRVHISTACTIVEENLARGE : BOOL
END_METHOD

(* ---- PROXYFBHISTALARMSROWQUEUE.pou ---- *)
FUNCTION_BLOCK PROXYFBHISTALARMSROWQUEUE
VAR
	M_PAHISTQUEUE : POINTER TO ARRAY [0..10] OF ProxyFbAlarmHistorical;
	M_ISZQUEUE : INT;
	MAXENTRIES : INT;
END_VAR
END_FUNCTION_BLOCK

METHOD FB_EXIT : BOOL
VAR_INPUT
	BINCOPYCODE : BOOL;
END_VAR
END_METHOD

METHOD GETAVAILABLEENTRIES : INT
END_METHOD

METHOD GETCOUNTTOREGISTER : INT
END_METHOD

METHOD GETITEM : POINTER TO ProxyFbAlarmHistorical
VAR_INPUT
	IOBJNUM : INT;
END_VAR
END_METHOD

METHOD INITIALIZE
VAR_INPUT
	SZQUEUE : INT;
END_VAR
END_METHOD

(* ---- REMOTEDEVICECOMPARER.pou ---- *)
FUNCTION_BLOCK REMOTEDEVICECOMPARER EXTENDS TSLastComparer
END_FUNCTION_BLOCK

METHOD COMPARE : INT
VAR_INPUT
	DIINDEXALARM1 : DINT;
	DIINDEXALARM2 : DINT;
END_VAR
END_METHOD

(* ---- REP_ACK_ALARMSTATEMACHINE.pou ---- *)
FUNCTION_BLOCK REP_ACK_ALARMSTATEMACHINE
END_FUNCTION_BLOCK

METHOD DOACKNOWLEDGE : AlarmState
VAR_INPUT
	ECURRENTSTATE : AlarmState;
END_VAR
VAR_OUTPUT
	ESTATETRANSITION : AlarmStateTransition;
END_VAR
END_METHOD

METHOD DOACTIVATE : AlarmState
VAR_INPUT
	ECURRENTSTATE : AlarmState;
END_VAR
END_METHOD

METHOD DODEACTIVATE : AlarmState
VAR_INPUT
	ECURRENTSTATE : AlarmState;
END_VAR
VAR_OUTPUT
	ESTATETRANSITION : AlarmStateTransition;
END_VAR
END_METHOD

(* ---- REP_ACK_ALARMSTATEMACHINE_NOCONFIRM.pou ---- *)
FUNCTION_BLOCK REP_ACK_ALARMSTATEMACHINE_NOCONFIRM EXTENDS Rep_Ack_AlarmStateMachine
END_FUNCTION_BLOCK

METHOD DOACKNOWLEDGE : AlarmState
VAR_INPUT
	ECURRENTSTATE : AlarmState;
END_VAR
VAR_OUTPUT
	ESTATETRANSITION : AlarmStateTransition;
END_VAR
END_METHOD

METHOD DODEACTIVATE : AlarmState
VAR_INPUT
	ECURRENTSTATE : AlarmState;
END_VAR
VAR_OUTPUT
	ESTATETRANSITION : AlarmStateTransition;
END_VAR
END_METHOD

(* ---- REP_ALARMSTATEMACHINE.pou ---- *)
FUNCTION_BLOCK REP_ALARMSTATEMACHINE
END_FUNCTION_BLOCK

METHOD DOACKNOWLEDGE : AlarmState
VAR_INPUT
	ECURRENTSTATE : AlarmState;
END_VAR
VAR_OUTPUT
	ESTATETRANSITION : AlarmStateTransition;
END_VAR
END_METHOD

METHOD DOACTIVATE : AlarmState
VAR_INPUT
	ECURRENTSTATE : AlarmState;
END_VAR
END_METHOD

METHOD DODEACTIVATE : AlarmState
VAR_INPUT
	ECURRENTSTATE : AlarmState;
END_VAR
VAR_OUTPUT
	ESTATETRANSITION : AlarmStateTransition;
END_VAR
END_METHOD

(* ---- REQUESTBUILDERACKALARMS.pou ---- *)
FUNCTION_BLOCK REQUESTBUILDERACKALARMS EXTENDS RequestBuilderBase
VAR
	M_ITFOWNSERVICEPROVIDER : IAckAlarmsServiceProvider;
	M_ITFOWNSERVICECONSUMER : IAckAlarmsServiceConsumer;
	COMPONENT : STRING := 'RequestBuilderReadActiveAlarms';
END_VAR
END_FUNCTION_BLOCK

METHOD BUILDANDENQUEUEV3REQUEST : UDINT
VAR_INPUT
	IREQUESTID : INT;
	ITFSERVICEPROVIDER : IServiceProvider;
	ITFSERVICECONSUMER : IServiceConsumer;
END_VAR
END_METHOD

METHOD FB_INIT : BOOL
VAR_INPUT
	BINITRETAINS : BOOL;
	BINCOPYCODE : BOOL;
END_VAR
END_METHOD

METHOD INITIALIZE
VAR_INPUT
	ITFDATASOURCE : IDatasources.IDatasource2;
	IMAXALMGROUPS : INT;
END_VAR
END_METHOD

METHOD BUILDREQUEST : UDINT
VAR_INPUT
	ITFSERVICEWRITER : CDSV3Prot.IServiceWriter;
	XHASTOSWAP : BOOL;
END_VAR
END_METHOD

METHOD GETSERVICE : UINT
END_METHOD

METHOD REQUESTFINISHED
VAR_INPUT
	REQUEST : IDatasources.ICustomRequest;
	RESPONSE : IDatasources.ICustomResponse;
	RESULT : SysTypes.RTS_IEC_RESULT;
END_VAR
END_METHOD

(* ---- REQUESTBUILDERBASE.pou ---- *)
FUNCTION_BLOCK REQUESTBUILDERBASE
VAR_INPUT
	M_REQUESTMONITOR : ProxyStructMonitorRequest;
	M_XLOCK : BOOL;
	M_HLOCK : RTS_IEC_HANDLE;
END_VAR
VAR
	M_ITFDATASOURCE : IDatasources.IDatasource2;
	M_ITFCDSV3REQUEST : IDatasources.ICDSV3Request;
	M_EBYTEORDER : IDatasources.ByteOrder := IDatasources.ByteOrder.Unknown;
	M_XHASTOSWAP : BOOL;
	M_ITFCDSV3REQUESTBUILDER : CDSV3Prot.ICDSV3RequestBuilder;
	M_ITFCUSTOMREQUESTCALLBACK : IDatasources.ICustomRequestCallback;
	M_PABYREQUESTBUFFER : POINTER TO BYTE;
	M_UDIREQUESTBUFFERSIZE : UDINT := MEM_SIZE_UNIT;
	M_ICURRREQUESTID : INT;
	M_IFBREQUESTID : INT;
	M_ITFSERVICECONSUMER : IServiceConsumer;
	M_LTSTARTTIME : LTIME;
	M_LTSTARTTIMEWAITANS : LTIME;
	M_UDIPREVERRCOUNT : UDINT;
	M_DURATION1 : Statistics_LTIME;
	M_IDURATIONSTATCNT : INT := 10;
	M_LTREQDURATIONLAST : LTIME;
	M_LTREQDURATIONAVG : LTIME;
	M_LTREQDURATIONMIN : LTIME;
	M_LTREQDURATIONMAX : LTIME;
	M_LTREQDURATIONBUILDREQ : LTIME;
	M_LTREQDURATIONWAITANS : LTIME;
	M_LTREQDURATIONELABANS : LTIME;
	M_SCOMPONENT : STRING := 'RequestBuilderBase';
	M_LOCKRESULT : RTS_IEC_RESULT := Errors.ERR_FAILED;
	MEM_SIZE_UNIT : UDINT := 256;
	MEM_SIZE_UNIT_GRP : UDINT := (MEM_SIZE_UNIT * 4);
	ISERRORPRESENT : BOOL;
END_VAR
END_FUNCTION_BLOCK

METHOD ADDERROR
VAR_INPUT
	UDIERROR : UDINT;
	SMSG : STRING;
END_VAR
END_METHOD

METHOD BUILDANDENQUEUEV3REQUEST : UDINT
VAR_INPUT
	IREQUESTID : INT;
	ITFSERVICEPROVIDER : IServiceProvider;
	ITFSERVICECONSUMER : IServiceConsumer;
END_VAR
END_METHOD

METHOD FB_EXIT : BOOL
VAR_INPUT
	BINCOPYCODE : BOOL;
END_VAR
END_METHOD

METHOD GETSTATISTICSDATA
END_METHOD

METHOD INITIALIZE
VAR_INPUT
	ITFDATASOURCE : IDatasources.IDatasource2;
	IMAXALMGROUPS : INT;
END_VAR
END_METHOD

METHOD BUILDREQUEST : UDINT
VAR_INPUT
	ITFSERVICEWRITER : CDSV3Prot.IServiceWriter;
	XHASTOSWAP : BOOL;
END_VAR
END_METHOD

METHOD GETDATABUFFER : POINTER TO BYTE
END_METHOD

METHOD GETDATABUFFERSIZE : UDINT
END_METHOD

METHOD GETSERVICE : UINT
END_METHOD

METHOD GETSERVICEGROUP : UINT
END_METHOD

METHOD REQUESTENQUEUED : UDINT
END_METHOD

METHOD SETTARGETBYTEORDER
VAR_INPUT
	EBYTEORDER : IDatasources.ByteOrder;
END_VAR
END_METHOD

METHOD REQUESTFINISHED
VAR_INPUT
	REQUEST : IDatasources.ICustomRequest;
	RESPONSE : IDatasources.ICustomResponse;
	RESULT : SysTypes.RTS_IEC_RESULT;
END_VAR
END_METHOD

METHOD PROTAFTERBUILDREQUEST
END_METHOD

METHOD PROTAFTERREQUEST
VAR_INPUT
	ITFSERVICECONSUMER : IServiceConsumer;
END_VAR
END_METHOD

METHOD PROTBEFOREANSELAB
END_METHOD

METHOD PROTBEFOREREQUEST
VAR_INPUT
	IREQUESTID : INT;
END_VAR
END_METHOD

METHOD PROTBUILDANDENQUEUEV3REQUEST : UDINT
END_METHOD

METHOD PROTRELEASEREQUEST
END_METHOD

(* ---- REQUESTBUILDERCHANNELTEST.pou ---- *)
FUNCTION_BLOCK REQUESTBUILDERCHANNELTEST EXTENDS RequestBuilderBase
VAR
	M_ITFOWNSERVICEPROVIDER : IChannelTestServiceProvider;
	M_ITFOWNSERVICECONSUMER : IChannelTestServiceConsumer;
	COMPONENT : STRING := 'RequestBuilderChannelTest';
END_VAR
END_FUNCTION_BLOCK

METHOD BUILDANDENQUEUEV3REQUEST : UDINT
VAR_INPUT
	IREQUESTID : INT;
	ITFSERVICEPROVIDER : IServiceProvider;
	ITFSERVICECONSUMER : IServiceConsumer;
END_VAR
END_METHOD

METHOD FB_INIT : BOOL
VAR_INPUT
	BINITRETAINS : BOOL;
	BINCOPYCODE : BOOL;
END_VAR
END_METHOD

METHOD INITIALIZE
VAR_INPUT
	ITFDATASOURCE : IDatasources.IDatasource2;
	IMAXALMGROUPS : INT;
END_VAR
END_METHOD

METHOD BUILDREQUEST : UDINT
VAR_INPUT
	ITFSERVICEWRITER : CDSV3Prot.IServiceWriter;
	XHASTOSWAP : BOOL;
END_VAR
END_METHOD

METHOD GETSERVICE : UINT
END_METHOD

METHOD REQUESTFINISHED
VAR_INPUT
	REQUEST : IDatasources.ICustomRequest;
	RESPONSE : IDatasources.ICustomResponse;
	RESULT : SysTypes.RTS_IEC_RESULT;
END_VAR
END_METHOD

(* ---- REQUESTBUILDERCHANNELTEST2.pou ---- *)
FUNCTION_BLOCK REQUESTBUILDERCHANNELTEST2 EXTENDS RequestBuilderChannelTest
VAR
	COMPONENT2 : STRING := 'RequestBuilderChannelTest2';
END_VAR
END_FUNCTION_BLOCK

METHOD FB_INIT : BOOL
VAR_INPUT
	BINITRETAINS : BOOL;
	BINCOPYCODE : BOOL;
END_VAR
END_METHOD

METHOD INITIALIZE
VAR_INPUT
	ITFDATASOURCE : IDatasources.IDatasource2;
	IMAXALMGROUPS : INT;
END_VAR
END_METHOD

(* ---- REQUESTBUILDERGETALMCLASSCONFIG.pou ---- *)
FUNCTION_BLOCK REQUESTBUILDERGETALMCLASSCONFIG EXTENDS RequestBuilderBase
VAR
	M_ITFOWNSERVICEPROVIDER : IAlmConfigServiceProvider;
	M_ITFOWNSERVICECONSUMER : IAlmConfigServiceConsumer;
	COMPONENT : STRING := 'RequestBuilderGetAlmClassConfig';
END_VAR
END_FUNCTION_BLOCK

METHOD BUILDANDENQUEUEV3REQUEST : UDINT
VAR_INPUT
	IREQUESTID : INT;
	ITFSERVICEPROVIDER : IServiceProvider;
	ITFSERVICECONSUMER : IServiceConsumer;
END_VAR
END_METHOD

METHOD FB_INIT : BOOL
VAR_INPUT
	BINITRETAINS : BOOL;
	BINCOPYCODE : BOOL;
END_VAR
END_METHOD

METHOD INITIALIZE
VAR_INPUT
	ITFDATASOURCE : IDatasources.IDatasource2;
	IMAXALMGROUPS : INT;
END_VAR
END_METHOD

METHOD BUILDREQUEST : UDINT
VAR_INPUT
	ITFSERVICEWRITER : CDSV3Prot.IServiceWriter;
	XHASTOSWAP : BOOL;
END_VAR
END_METHOD

METHOD GETSERVICE : UINT
END_METHOD

METHOD REQUESTFINISHED
VAR_INPUT
	REQUEST : IDatasources.ICustomRequest;
	RESPONSE : IDatasources.ICustomResponse;
	RESULT : SysTypes.RTS_IEC_RESULT;
END_VAR
END_METHOD

(* ---- REQUESTBUILDERGETALMCONFIG.pou ---- *)
FUNCTION_BLOCK REQUESTBUILDERGETALMCONFIG EXTENDS RequestBuilderBase
VAR
	M_ITFOWNSERVICEPROVIDER : IAlmConfigServiceProvider;
	M_ITFOWNSERVICECONSUMER : IAlmConfigServiceConsumer;
	COMPONENT : STRING := 'RequestBuilderGetAlmConfig';
END_VAR
END_FUNCTION_BLOCK

METHOD BUILDANDENQUEUEV3REQUEST : UDINT
VAR_INPUT
	IREQUESTID : INT;
	ITFSERVICEPROVIDER : IServiceProvider;
	ITFSERVICECONSUMER : IServiceConsumer;
END_VAR
END_METHOD

METHOD FB_INIT : BOOL
VAR_INPUT
	BINITRETAINS : BOOL;
	BINCOPYCODE : BOOL;
END_VAR
END_METHOD

METHOD INITIALIZE
VAR_INPUT
	ITFDATASOURCE : IDatasources.IDatasource2;
	IMAXALMGROUPS : INT;
END_VAR
END_METHOD

METHOD BUILDREQUEST : UDINT
VAR_INPUT
	ITFSERVICEWRITER : CDSV3Prot.IServiceWriter;
	XHASTOSWAP : BOOL;
END_VAR
END_METHOD

METHOD GETSERVICE : UINT
END_METHOD

METHOD REQUESTFINISHED
VAR_INPUT
	REQUEST : IDatasources.ICustomRequest;
	RESPONSE : IDatasources.ICustomResponse;
	RESULT : SysTypes.RTS_IEC_RESULT;
END_VAR
END_METHOD

(* ---- REQUESTBUILDERGETHISTORICALALMCONFIG.pou ---- *)
FUNCTION_BLOCK REQUESTBUILDERGETHISTORICALALMCONFIG EXTENDS RequestBuilderBase
VAR
	M_ITFOWNSERVICEPROVIDER : IHistoricAlmServiceProvider;
	M_ITFOWNSERVICECONSUMER : IHistoricAlmServiceConsumer;
	COMPONENT : STRING := 'RequestBuilderGetHistoricalAlmConfig';
END_VAR
END_FUNCTION_BLOCK

METHOD BUILDANDENQUEUEV3REQUEST : UDINT
VAR_INPUT
	IREQUESTID : INT;
	ITFSERVICEPROVIDER : IServiceProvider;
	ITFSERVICECONSUMER : IServiceConsumer;
END_VAR
END_METHOD

METHOD FB_INIT : BOOL
VAR_INPUT
	BINITRETAINS : BOOL;
	BINCOPYCODE : BOOL;
END_VAR
END_METHOD

METHOD INITIALIZE
VAR_INPUT
	ITFDATASOURCE : IDatasources.IDatasource2;
	IMAXALMGROUPS : INT;
END_VAR
END_METHOD

METHOD BUILDREQUEST : UDINT
VAR_INPUT
	ITFSERVICEWRITER : CDSV3Prot.IServiceWriter;
	XHASTOSWAP : BOOL;
END_VAR
END_METHOD

METHOD GETSERVICE : UINT
END_METHOD

METHOD REQUESTFINISHED
VAR_INPUT
	REQUEST : IDatasources.ICustomRequest;
	RESPONSE : IDatasources.ICustomResponse;
	RESULT : SysTypes.RTS_IEC_RESULT;
END_VAR
END_METHOD

(* ---- REQUESTBUILDERREADACTIVEALARMS.pou ---- *)
FUNCTION_BLOCK REQUESTBUILDERREADACTIVEALARMS EXTENDS RequestBuilderBase
VAR
	M_ITFOWNSERVICEPROVIDER : IReadActiveAlarmsServiceProvider;
	M_ITFOWNSERVICECONSUMER : IReadActiveAlarmsServiceConsumer;
	COMPONENT : STRING := 'RequestBuilderReadActiveAlarms';
END_VAR
END_FUNCTION_BLOCK

METHOD BUILDANDENQUEUEV3REQUEST : UDINT
VAR_INPUT
	IREQUESTID : INT;
	ITFSERVICEPROVIDER : IServiceProvider;
	ITFSERVICECONSUMER : IServiceConsumer;
END_VAR
END_METHOD

METHOD FB_INIT : BOOL
VAR_INPUT
	BINITRETAINS : BOOL;
	BINCOPYCODE : BOOL;
END_VAR
END_METHOD

METHOD INITIALIZE
VAR_INPUT
	ITFDATASOURCE : IDatasources.IDatasource2;
	IMAXALMGROUPS : INT;
END_VAR
END_METHOD

METHOD BUILDREQUEST : UDINT
VAR_INPUT
	ITFSERVICEWRITER : CDSV3Prot.IServiceWriter;
	XHASTOSWAP : BOOL;
END_VAR
END_METHOD

METHOD GETSERVICE : UINT
END_METHOD

METHOD REQUESTFINISHED
VAR_INPUT
	REQUEST : IDatasources.ICustomRequest;
	RESPONSE : IDatasources.ICustomResponse;
	RESULT : SysTypes.RTS_IEC_RESULT;
END_VAR
END_METHOD

(* ---- REQUESTBUILDERREADHISTORICALACTIVEALARMS.pou ---- *)
FUNCTION_BLOCK REQUESTBUILDERREADHISTORICALACTIVEALARMS EXTENDS RequestBuilderBase
VAR
	M_ITFOWNSERVICEPROVIDER : IHistoricAlmServiceProvider;
	M_ITFOWNSERVICECONSUMER : IHistoricAlmServiceConsumer;
	COMPONENT : STRING := 'RequestBuilderReadHistoricalActiveAlarms';
END_VAR
END_FUNCTION_BLOCK

METHOD BUILDANDENQUEUEV3REQUEST : UDINT
VAR_INPUT
	IREQUESTID : INT;
	ITFSERVICEPROVIDER : IServiceProvider;
	ITFSERVICECONSUMER : IServiceConsumer;
END_VAR
END_METHOD

METHOD FB_INIT : BOOL
VAR_INPUT
	BINITRETAINS : BOOL;
	BINCOPYCODE : BOOL;
END_VAR
END_METHOD

METHOD INITIALIZE
VAR_INPUT
	ITFDATASOURCE : IDatasources.IDatasource2;
	IMAXALMGROUPS : INT;
END_VAR
END_METHOD

METHOD BUILDREQUEST : UDINT
VAR_INPUT
	ITFSERVICEWRITER : CDSV3Prot.IServiceWriter;
	XHASTOSWAP : BOOL;
END_VAR
END_METHOD

METHOD GETSERVICE : UINT
END_METHOD

METHOD REQUESTFINISHED
VAR_INPUT
	REQUEST : IDatasources.ICustomRequest;
	RESPONSE : IDatasources.ICustomResponse;
	RESULT : SysTypes.RTS_IEC_RESULT;
END_VAR
END_METHOD

(* ---- REQUESTBUILDERREADHISTORICALALARMS.pou ---- *)
FUNCTION_BLOCK REQUESTBUILDERREADHISTORICALALARMS EXTENDS RequestBuilderBase
VAR
	M_ITFOWNSERVICEPROVIDER : IHistoricAlmServiceProvider;
	M_ITFOWNSERVICECONSUMER : IHistoricAlmServiceConsumer;
	COMPONENT : STRING := 'RequestBuilderReadHistoricalAlarms';
END_VAR
END_FUNCTION_BLOCK

METHOD BUILDANDENQUEUEV3REQUEST : UDINT
VAR_INPUT
	IREQUESTID : INT;
	ITFSERVICEPROVIDER : IServiceProvider;
	ITFSERVICECONSUMER : IServiceConsumer;
END_VAR
END_METHOD

METHOD FB_INIT : BOOL
VAR_INPUT
	BINITRETAINS : BOOL;
	BINCOPYCODE : BOOL;
END_VAR
END_METHOD

METHOD INITIALIZE
VAR_INPUT
	ITFDATASOURCE : IDatasources.IDatasource2;
	IMAXALMGROUPS : INT;
END_VAR
END_METHOD

METHOD BUILDREQUEST : UDINT
VAR_INPUT
	ITFSERVICEWRITER : CDSV3Prot.IServiceWriter;
	XHASTOSWAP : BOOL;
END_VAR
END_METHOD

METHOD GETSERVICE : UINT
END_METHOD

METHOD REQUESTFINISHED
VAR_INPUT
	REQUEST : IDatasources.ICustomRequest;
	RESPONSE : IDatasources.ICustomResponse;
	RESULT : SysTypes.RTS_IEC_RESULT;
END_VAR
END_METHOD

(* ---- REQUESTBUILDERRESETALMRECORD.pou ---- *)
FUNCTION_BLOCK REQUESTBUILDERRESETALMRECORD EXTENDS RequestBuilderBase
VAR
	M_ITFOWNSERVICEPROVIDER : IAlmRecordServiceProvider;
	M_ITFOWNSERVICECONSUMER : IAlmRecordServiceConsumer;
	COMPONENT : STRING := 'RequestBuilderResetAlmRecord';
END_VAR
END_FUNCTION_BLOCK

METHOD BUILDANDENQUEUEV3REQUEST : UDINT
VAR_INPUT
	IREQUESTID : INT;
	ITFSERVICEPROVIDER : IServiceProvider;
	ITFSERVICECONSUMER : IServiceConsumer;
END_VAR
END_METHOD

METHOD FB_INIT : BOOL
VAR_INPUT
	BINITRETAINS : BOOL;
	BINCOPYCODE : BOOL;
END_VAR
END_METHOD

METHOD INITIALIZE
VAR_INPUT
	ITFDATASOURCE : IDatasources.IDatasource2;
	IMAXALMGROUPS : INT;
END_VAR
END_METHOD

METHOD BUILDREQUEST : UDINT
VAR_INPUT
	ITFSERVICEWRITER : CDSV3Prot.IServiceWriter;
	XHASTOSWAP : BOOL;
END_VAR
END_METHOD

METHOD GETSERVICE : UINT
END_METHOD

METHOD REQUESTFINISHED
VAR_INPUT
	REQUEST : IDatasources.ICustomRequest;
	RESPONSE : IDatasources.ICustomResponse;
	RESULT : SysTypes.RTS_IEC_RESULT;
END_VAR
END_METHOD

(* ---- REQUESTBUILDERSETALMRECORD.pou ---- *)
FUNCTION_BLOCK REQUESTBUILDERSETALMRECORD EXTENDS RequestBuilderBase
VAR
	M_ITFOWNSERVICEPROVIDER : IAlmRecordServiceProvider;
	M_ITFOWNSERVICECONSUMER : IAlmRecordServiceConsumer;
	COMPONENT : STRING := 'RequestBuilderSetAlmRecord';
END_VAR
END_FUNCTION_BLOCK

METHOD BUILDANDENQUEUEV3REQUEST : UDINT
VAR_INPUT
	IREQUESTID : INT;
	ITFSERVICEPROVIDER : IServiceProvider;
	ITFSERVICECONSUMER : IServiceConsumer;
END_VAR
END_METHOD

METHOD FB_INIT : BOOL
VAR_INPUT
	BINITRETAINS : BOOL;
	BINCOPYCODE : BOOL;
END_VAR
END_METHOD

METHOD INITIALIZE
VAR_INPUT
	ITFDATASOURCE : IDatasources.IDatasource2;
	IMAXALMGROUPS : INT;
END_VAR
END_METHOD

METHOD BUILDREQUEST : UDINT
VAR_INPUT
	ITFSERVICEWRITER : CDSV3Prot.IServiceWriter;
	XHASTOSWAP : BOOL;
END_VAR
END_METHOD

METHOD GETSERVICE : UINT
END_METHOD

METHOD REQUESTFINISHED
VAR_INPUT
	REQUEST : IDatasources.ICustomRequest;
	RESPONSE : IDatasources.ICustomResponse;
	RESULT : SysTypes.RTS_IEC_RESULT;
END_VAR
END_METHOD

(* ---- ROWIDCOMPARER.pou ---- *)
FUNCTION_BLOCK ROWIDCOMPARER EXTENDS AbstractComparer
END_FUNCTION_BLOCK

METHOD COMPARE : INT
VAR_INPUT
	DIINDEXALARM1 : DINT;
	DIINDEXALARM2 : DINT;
END_VAR
END_METHOD

(* ---- RUNTIMEEVENTLISTENER.pou ---- *)
FUNCTION_BLOCK RUNTIMEEVENTLISTENER
VAR
	_HPREPAREDOWNLOADEVENT : RTS_IEC_HANDLE := Events.Invalid_Handle;
	_HPREPAREDOWNLOADEVENTINTERFACE : RTS_IEC_HANDLE := Events.Invalid_Handle;
	_HPREPARESTOPEVENT : RTS_IEC_HANDLE := Events.Invalid_Handle;
	_HPREPARESTOPEVENTINTERFACE : RTS_IEC_HANDLE := Events.Invalid_Handle;
END_VAR
END_FUNCTION_BLOCK

METHOD EVENTCALLBACK : UDINT
VAR_INPUT
	PEVENTPARAM : POINTER TO EventParam;
END_VAR
END_METHOD

METHOD FB_EXIT : BOOL
VAR_INPUT
	BINCOPYCODE : BOOL;
END_VAR
END_METHOD

METHOD FB_INIT : BOOL
VAR_INPUT
	BINITRETAINS : BOOL;
	BINCOPYCODE : BOOL;
END_VAR
END_METHOD

METHOD PRVISOURAPPLICATIONBEFOREDELETE : BOOL
VAR_INPUT
	PAPPDELETEEVENTPARAM : POINTER TO CmPApp.EVTPARAM_CmpAppStop;
END_VAR
END_METHOD

METHOD PRVISOURAPPLICATIONBEFOREDOWNLOAD : BOOL
VAR_INPUT
	PAPPEVENTPARAM : POINTER TO CmPApp.EVTPARAM_CmpApp;
END_VAR
END_METHOD

(* ---- SERIALIZERDATABLOCK.pou ---- *)
FUNCTION_BLOCK SERIALIZERDATABLOCK
VAR_INPUT
	M_PBYBUFFER : POINTER TO BYTE;
	M_UDIBUFFERSIZE : UDINT;
END_VAR
VAR
	M_SERIALIZINGALARMMETAOBJECTSTUB : SerializingAlarmMetaObjectStub;
	M_ICOUNTROWS : INT;
	ERROR : UINT;
END_VAR
END_FUNCTION_BLOCK

METHOD GETALARMMETAOBJECTSTUB : IAlarmMetaObjectStub3
VAR_INPUT
	IROW : INT;
	IOFFSET : INT;
END_VAR
END_METHOD

METHOD GETCOUNTROWS : INT
END_METHOD

METHOD SETCOUNTROWS : BOOL
VAR_INPUT
	ICOUNT : INT;
END_VAR
END_METHOD

METHOD HASALARMS : BOOL
END_METHOD

METHOD SETTOTALCOUNTROWS : BOOL
VAR_INPUT
	DICOUNT : DINT;
END_VAR
END_METHOD

(* ---- SERIALIZINGALARMMETAOBJECTSTUB.pou ---- *)
FUNCTION_BLOCK SERIALIZINGALARMMETAOBJECTSTUB
VAR_INPUT
	M_PBYBUFFER : POINTER TO BYTE;
	M_UDIBUFFERSIZE : UDINT;
	M_UDIOFFSET : UDINT;
	M_XOVERFLOW : BOOL;
END_VAR
VAR
	S_OFFSET_TIMESTAMP_LAST : UDINT := 0;
	S_OFFSET_TIMESTAMP_ACTIVE : UDINT := (8 + s_OFFSET_TIMESTAMP_LAST);
	S_OFFSET_TIMESTAMP_INACTIVE : UDINT := (8 + s_OFFSET_TIMESTAMP_ACTIVE);
	S_OFFSET_TIMESTAMP_ACKNOWLEDGE : UDINT := (8 + s_OFFSET_TIMESTAMP_INACTIVE);
	S_OFFSET_TRIGGER_VALUE : UDINT := (8 + s_OFFSET_TIMESTAMP_ACKNOWLEDGE);
	S_OFFSET_LATCH1_VALUE : UDINT := (8 + s_OFFSET_TRIGGER_VALUE);
	S_OFFSET_LATCH2_VALUE : UDINT := (8 + s_OFFSET_LATCH1_VALUE);
	S_OFFSET_ALARMGROUP_ID : UDINT := (8 + s_OFFSET_LATCH2_VALUE);
	S_OFFSET_ALARM_ID : UDINT := (4 + s_OFFSET_ALARMGROUP_ID);
	S_OFFSET_STATE : UDINT := (4 + s_OFFSET_ALARM_ID);
	S_OFFSET_TRIGGER_VALUE_TYPE : UDINT := (1 + s_OFFSET_STATE);
	S_OFFSET_LATCH1_TYPE : UDINT := (1 + s_OFFSET_TRIGGER_VALUE_TYPE);
	S_OFFSET_LATCH2_TYPE : UDINT := (1 + s_OFFSET_LATCH1_TYPE);
	SIZE_LATCH2_TYPE : UDINT := 1;
	SIZE : UDINT;
END_VAR
END_FUNCTION_BLOCK

METHOD INITIALIZE
END_METHOD

METHOD SETALARM
VAR_INPUT
	PALARM : POINTER TO Alarm;
END_VAR
END_METHOD

METHOD SETLATCHVAR1VALUE
VAR_INPUT
	ITFTYPEDVALUELATCHVAR1 : ITypedValue;
END_VAR
END_METHOD

METHOD SETLATCHVAR2VALUE
VAR_INPUT
	ITFTYPEDVALUELATCHVAR2 : ITypedValue;
END_VAR
END_METHOD

METHOD SETSTATE
VAR_INPUT
	ISTATE : INT;
END_VAR
END_METHOD

METHOD SETTIMESTAMPACKNOWLEDGE
VAR_INPUT
	LITIMESTAMPACKNOWLEDGE : Timestamp;
END_VAR
END_METHOD

METHOD SETTIMESTAMPACTIVE
VAR_INPUT
	LITIMESTAMPACTIVE : Timestamp;
END_VAR
END_METHOD

METHOD SETTIMESTAMPINACTIVE
VAR_INPUT
	LITIMESTAMPINACTIVE : Timestamp;
END_VAR
END_METHOD

METHOD SETTIMESTAMPLAST
VAR_INPUT
	LITIMESTAMPLAST : Timestamp;
END_VAR
END_METHOD

METHOD SETTRIGGERVALUE
VAR_INPUT
	ITFTYPEDVALUETRIGGER : ITypedValue;
END_VAR
END_METHOD

METHOD GETALARM : POINTER TO Alarm
END_METHOD

METHOD GETALARMGROUP : STRING
END_METHOD

METHOD GETCHECKSUM : UDINT
END_METHOD

METHOD GETCURRENTVALUE : ITypedValue
END_METHOD

METHOD GETID : ALARM_ID
END_METHOD

METHOD GETLATCHVAR1VALUE : ITypedValue
END_METHOD

METHOD GETLATCHVAR2VALUE : ITypedValue
END_METHOD

METHOD GETSTATE : INT
END_METHOD

METHOD GETTIMESTAMPACKNOWLEDGE : Timestamp
END_METHOD

METHOD GETTIMESTAMPACTIVE : Timestamp
END_METHOD

METHOD GETTIMESTAMPINACTIVE : Timestamp
END_METHOD

METHOD GETTIMESTAMPLAST : Timestamp
END_METHOD

METHOD GETTRIGGERVALUE : ITypedValue
END_METHOD

METHOD SETACKNOWLEDGE
VAR_INPUT
	BACKNOWLEDGEMULTIPLE : BOOL;
END_VAR
END_METHOD

METHOD SETALARMGROUP
VAR_INPUT
	SALARMGROUP : STRING;
END_VAR
END_METHOD

METHOD SETCURRENTLREALVALUE
VAR_INPUT
	LRVALUE : LREAL;
END_VAR
END_METHOD

METHOD SETCURRENTVALUE
VAR_INPUT
	ITFTYPEDVALUECURRENT : ITypedValue;
END_VAR
END_METHOD

METHOD SETID
VAR_INPUT
	UIID : ALARM_ID;
END_VAR
END_METHOD

(* ---- SQLITEDATABASEACCESS.pou ---- *)
FUNCTION_BLOCK SQLITEDATABASEACCESS EXTENDS AbstractDatabaseAccess
VAR
	M_CONTEXT : SQLiteDatabaseAccessContext;
	M_ITFALARMSTORAGEMANAGER : IAlarmStorageManager;
	M_ISUPPORTEDVERSION : INT := -1;
	M_XBYTEORDERGET : BOOL;
END_VAR
END_FUNCTION_BLOCK

METHOD SETALARMSTORAGEMANAGER
VAR_INPUT
	ITFALARMSTORAGEMANAGER : IAlarmStorageManager;
END_VAR
END_METHOD

METHOD GETNUMBEROFLATCHVARIABLES : USINT
END_METHOD

METHOD GETROOTPAGE : CAA.IDENT
VAR_INPUT
	EWHICHALARMSTORAGEOBJECT : EAlarmStorageObject;
END_VAR
END_METHOD

METHOD ISONLYONEALARMCLASSSELECTED : BOOL
END_METHOD

METHOD ISONLYONEALARMGROUPSELECTED : BOOL
END_METHOD

METHOD PREPAREDATABASEACCESS : STO.ERROR
END_METHOD

METHOD TBLALARMCURSORCLOSE : STO.ERROR
VAR_INPUT
	EERRORFROMPREVIOUSPROCESSING : STO.ERROR;
END_VAR
END_METHOD

METHOD TBLALARMCURSORMOVE : STO.ERROR
VAR_INPUT
	EDIRECTION : STO.DIRECTION;
END_VAR
VAR_OUTPUT
	XEOF : BOOL;
END_VAR
END_METHOD

METHOD TBLALARMCURSOROPEN : STO.ERROR
VAR_INPUT
	FILTERCRITERIA : REFERENCE TO VisuFbAlarmFilterCriteria;
END_VAR
END_METHOD

METHOD TBLALARMCURSOROPEN2 : STO.ERROR
VAR_INPUT
	IDINDEX : CAA.IDENT;
END_VAR
END_METHOD

METHOD TBLALARMCURSORSETPOSITION : STO.ERROR
VAR_INPUT
	FILTERCRITERIA : REFERENCE TO VisuFbAlarmFilterCriteria;
	BROWIDVALID : BOOL;
	DIROWID : DINT;
END_VAR
END_METHOD

METHOD TBLALARMGETLATCHVARTYPE : STO.ERROR
VAR_INPUT
	IDWHICHCOLUMN : CAA.IDENT;
	USIWHICHLATCHVAR : USINT;
END_VAR
VAR_OUTPUT
	BYTYPE : BYTE;
	XNULL : BOOL;
END_VAR
END_METHOD

METHOD TBLALARMGETLATCHVARVALUE : STO.ERROR
VAR_INPUT
	IDWHICHCOLUMN : CAA.IDENT;
	USIWHICHLATCHVAR : USINT;
END_VAR
VAR_OUTPUT
	LIVALUE : LINT;
	XNULL : BOOL;
END_VAR
END_METHOD

METHOD TBLALARMGETMINMAXROWIDS : BOOL
VAR_OUTPUT
	IDROWMIN : LINT;
	IDROWMAX : LINT;
	EERROR : STO.ERROR;
END_VAR
END_METHOD

METHOD TBLALARMGETROWCOUNT : CAA.COUNT
VAR_OUTPUT
	EERROR : STO.ERROR;
END_VAR
END_METHOD

METHOD TBLALARMGETTIMESTAMPVALUE : LINT
VAR_INPUT
	IDWHICHCOLUMN : CAA.IDENT;
END_VAR
VAR_OUTPUT
	EERROR : STO.ERROR;
END_VAR
END_METHOD

METHOD TBLALARMGET_DINT : STO.ERROR
VAR_INPUT
	IDWHICHCOLUMN : CAA.IDENT;
	IWHICHCOLUMN : INT;
END_VAR
VAR_OUTPUT
	DIVALUE : DINT;
	XNULL : BOOL;
END_VAR
END_METHOD

METHOD TBLALARMGET_LINT : STO.ERROR
VAR_INPUT
	IDWHICHCOLUMN : CAA.IDENT;
	IWHICHCOLUMN : INT;
END_VAR
VAR_OUTPUT
	LIVALUE : LINT;
	XNULL : BOOL;
END_VAR
END_METHOD

METHOD TBLALARMGET_SINT : STO.ERROR
VAR_INPUT
	IDWHICHCOLUMN : CAA.IDENT;
	IWHICHCOLUMN : INT;
END_VAR
VAR_OUTPUT
	SIVALUE : SINT;
	XNULL : BOOL;
END_VAR
END_METHOD

METHOD TBLALARMISNOTEMPTY : BOOL
VAR_OUTPUT
	EERROR : STO.ERROR;
END_VAR
END_METHOD

METHOD TBLALARMROWGETCURRENT : STO.ERROR
END_METHOD

METHOD TBLALARMROWGETCURRENTID : DINT
END_METHOD

METHOD TBLALARMROWISVALID : BOOL
END_METHOD

METHOD TBLALARMROWRELEASE : STO.ERROR
VAR_INPUT
	EERRORFROMPREVIOUSPROCESSING : STO.ERROR;
END_VAR
END_METHOD

METHOD TBLALARMROWSELECT : STO.ERROR
VAR_INPUT
	IDROW : CAA.IDENT;
	XDOERRORHANDLING : BOOL;
END_VAR
END_METHOD

METHOD TBLALARMTABLECLOSE : STO.ERROR
END_METHOD

METHOD TBLALARMTABLEISOPEN : BOOL
END_METHOD

METHOD TBLALARMTABLEOPEN : STO.ERROR
VAR_INPUT
	XREADONLY : BOOL;
END_VAR
END_METHOD

METHOD TBLLATCHVARSTRINGSCLOSEIFNEEDED : STO.ERROR
VAR_INPUT
	EERRORFROMPREVIOUSPROCESSING : STO.ERROR;
END_VAR
END_METHOD

METHOD TBLLATCHVARSTRINGSCURSORSEARCHROWID : STO.ERROR
VAR_INPUT
	LIROWID : LINT;
END_VAR
END_METHOD

METHOD TBLLATCHVARSTRINGSGET_TEXT : STO.ERROR
VAR_INPUT
	IDWHICHCOLUMN : CAA.IDENT;
	IWHICHCOLUMN : INT;
END_VAR
VAR_OUTPUT
	XNULL : BOOL;
END_VAR
VAR_IN_OUT
	TXTVALUE : STO.TEXT;
END_VAR
END_METHOD

METHOD TBLLATCHVARSTRINGSOPENIFNEEDED : STO.ERROR
END_METHOD

METHOD TBLLATCHVARSTRINGSROWGETCURRENT : STO.ERROR
END_METHOD

METHOD TBLLATCHVARSTRINGSROWRELEASE : STO.ERROR
VAR_INPUT
	EERRORFROMPREVIOUSPROCESSING : STO.ERROR;
END_VAR
END_METHOD

METHOD TEXTCOPYTOSTRING : STO.ERROR
VAR_INPUT
	XFREE : BOOL;
END_VAR
VAR_IN_OUT
	TXTVALUE : STO.TEXT;
	SVALUE : STRING(1);
	SZVALUE : CAA.SIZE;
END_VAR
END_METHOD

METHOD TEXTCOPYTOWSTRING : STO.ERROR
VAR_INPUT
	XFREE : BOOL;
END_VAR
VAR_IN_OUT
	TXTVALUE : STO.TEXT;
	WSVALUE : WSTRING(1);
	SZVALUE : CAA.SIZE;
END_VAR
END_METHOD

METHOD TRANSACTIONBEGIN : STO.ERROR
VAR_INPUT
	XREADONLY : BOOL;
END_VAR
END_METHOD

METHOD TRANSACTIONBEGINFAILED : BOOL
END_METHOD

METHOD TRANSACTIONEND
VAR_INPUT
	EERRORFROMPREVIOUSPROCESSING : STO.ERROR;
END_VAR
END_METHOD

METHOD TBLALARMGET_INT : STO.ERROR
VAR_INPUT
	IDWHICHCOLUMN : CAA.IDENT;
	IWHICHCOLUMN : INT;
END_VAR
VAR_OUTPUT
	IVALUE : INT;
	XNULL : BOOL;
END_VAR
END_METHOD

METHOD TBLVERSIONGETCURRENT : STO.ERROR
VAR_OUTPUT
	IVERSION : INT;
END_VAR
END_METHOD

METHOD GETRELEVANTFILTERDATA
VAR_OUTPUT
	EDBBYTEORDER : EAlarmByteOrder;
END_VAR
END_METHOD

METHOD TBLALARMCURSORSEARCHROWID : STO.ERROR
VAR_INPUT
	IDROW : DINT;
END_VAR
END_METHOD

METHOD TBLGETBYTEORDER : STO.ERROR
VAR_OUTPUT
	EBYTEORDER : EAlarmByteOrder;
END_VAR
END_METHOD

METHOD TBLVERSIONGETCURRENT2 : STO.ERROR
VAR_OUTPUT
	IVERSION : INT;
	EDBUSED : EDBType;
END_VAR
END_METHOD

METHOD TBLALARMGETCOMMENTVALUE : STO.ERROR
VAR_INPUT
	IDWHICHCOLUMN : CAA.IDENT;
	IWHICHCOLUMN : INT;
END_VAR
VAR_OUTPUT
	XNULL : BOOL;
END_VAR
VAR_IN_OUT
	WSVALUE : WSTRING(2000);
END_VAR
END_METHOD
